// TIA Portal V19 program export: 0 tag tables, 0 data types, 8 data blocks, 41 code blocks (in call order from the OBs), 0 instance data blocks

DATA_BLOCK "ROLL_DB15"   // DB4
{ S7_Optimized_Access := 'TRUE' }
VERSION : 0.1
// stored: AutoNumber true, DBAccessibleFromOPCUA true, DBAccessibleFromWebserver true, IsOnlyStoredInLoadMemory false, IsRetainMemResEnabled false, IsWriteProtectedInAS false, MemoryReserve 100
   VAR RETAIN
      DW : Array[0..131] of Word;
   END_VAR
BEGIN
   DW[0..16] := WORD#16#FFFF;
   DW[17] := WORD#16#3360;
   DW[18..23] := WORD#16#FFFF;
   DW[24] := WORD#16#1010;
   DW[25] := WORD#16#1020;
   DW[26..30] := WORD#16#FFFF;
   DW[31..32] := WORD#16#3120;
   DW[33] := WORD#16#2900;
   DW[34..52] := WORD#16#FFFF;
   DW[53..54] := WORD#16#2120;
   DW[55] := WORD#16#1010;
   DW[56] := WORD#16#2060;
   DW[57] := WORD#16#FFFF;
   DW[58..59] := WORD#16#3180;
   DW[60] := WORD#16#2060;
   DW[61..62] := WORD#16#2600;
   DW[63] := WORD#16#2010;
   DW[64] := WORD#16#FFFF;
   DW[65] := WORD#16#2015;
   DW[66] := WORD#16#FFFF;
   DW[67] := WORD#16#1050;
   DW[68..74] := WORD#16#FFFF;
   DW[75] := WORD#16#2600;
   DW[76] := WORD#16#FFFF;
   DW[77] := WORD#16#2300;
   DW[78..84] := WORD#16#FFFF;
   DW[85] := WORD#16#2120;
   DW[86..101] := WORD#16#FFFF;
   DW[102..103] := WORD#16#2300;
   DW[104..105] := WORD#16#FFFF;
   DW[106] := WORD#16#2010;
   DW[107] := WORD#16#2015;
   DW[108..114] := WORD#16#FFFF;
   DW[115..117] := WORD#16#1050;
   DW[118..126] := WORD#16#FFFF;
   DW[127] := WORD#16#0038;
   DW[128..129] := WORD#16#0011;
   DW[130] := WORD#16#3360;
END_DATA_BLOCK

DATA_BLOCK "ROLL_DB19"   // DB5
{ S7_Optimized_Access := 'TRUE' }
VERSION : 0.1
// stored: AutoNumber true, DBAccessibleFromOPCUA true, DBAccessibleFromWebserver true, IsOnlyStoredInLoadMemory false, IsRetainMemResEnabled false, IsWriteProtectedInAS false, MemoryReserve 100
   VAR RETAIN
      DW : Array[0..131] of Word;
   END_VAR
BEGIN
   DW[0] := WORD#16#FFFF;
   DW[1] := WORD#16#0020;
   DW[2] := WORD#16#0014;
   DW[3..127] := WORD#16#FFFF;
   DW[128..129] := WORD#16#0001;
   DW[130] := WORD#16#0020;
END_DATA_BLOCK

DATA_BLOCK "ROLL_DB205"   // DB8
{ S7_Optimized_Access := 'TRUE' }
VERSION : 0.1
// stored: AutoNumber true, DBAccessibleFromOPCUA true, DBAccessibleFromWebserver true, IsOnlyStoredInLoadMemory false, IsRetainMemResEnabled false, IsWriteProtectedInAS false, MemoryReserve 100
   VAR RETAIN
      DW : Array[0..41] of Word;
   END_VAR
BEGIN
   DW[5] := WORD#16#2360;
   DW[9] := WORD#16#2090;
   DW[13] := WORD#16#0001;
   DW[17] := WORD#16#2240;
   DW[21] := WORD#16#2060;
   DW[25] := WORD#16#2300;
   DW[29] := WORD#16#2120;
   DW[33] := WORD#16#2400;
   DW[37] := WORD#16#0001;
END_DATA_BLOCK

DATA_BLOCK "ROLL_HMI"   // DB3
{ S7_Optimized_Access := 'TRUE' }
VERSION : 0.1
// Flat, symbolic WinCC interface; TP900 control binding is a separate build step.
// stored: AutoNumber true, DBAccessibleFromOPCUA true, DBAccessibleFromWebserver true, IsOnlyStoredInLoadMemory false, IsRetainMemResEnabled false, IsWriteProtectedInAS false, MemoryReserve 100
   VAR
      Heartbeat : DInt;
      Connected : Bool;
      ManualFunction : Int := 255;
      GroundHeld : Bool;
      WorkHeld : Bool;
      KeyF : Array[1..16] of Bool;
      SelectedProgram : Int := 1;
      RecipeCommand : Int := 1;
      RecipeRequest : DInt;
      RecipeAck : DInt;
      RecipeError : Int;
      CurrentProgram : Int := 1;
      ParameterRequest : DInt;
      ParameterAck : DInt;
      ParameterDb : Int := 15;
      ParameterIndex : Int;
      ParameterValue : DInt;
      ParameterCurrentValue : DInt;
      ParameterSlotPresent : Bool;
      ParameterError : Int;
      Dwell1Seconds : Int := 360;
      Drain1Seconds : Int := 90;
      Ultrasound1 : Bool := TRUE;
      Dwell2Seconds : Int := 240;
      Drain2Seconds : Int := 60;
      Dwell3Seconds : Int := 300;
      Drain3Seconds : Int := 120;
      Dry4Seconds : Int := 400;
      BasketMotion : Int := 1;
      BathLift : Bool;
      ProcessTimer1Units : Int;
      ProcessTimer2Units : Int;
      StatusM : Array[0..255, 0..7] of Bool;
      LogicalOutputs : Array[16..25, 0..7] of Bool;
   END_VAR
BEGIN
END_DATA_BLOCK

DATA_BLOCK "ROLL_IO"   // DB2
{ S7_Optimized_Access := 'TRUE' }
VERSION : 0.1
// stored: AutoNumber true, DBAccessibleFromOPCUA true, DBAccessibleFromWebserver true, IsOnlyStoredInLoadMemory false, IsRetainMemResEnabled false, IsWriteProtectedInAS false, MemoryReserve 100
   VAR
      Input : Array[0..127, 0..7] of Bool;
      Output : Array[0..127, 0..7] of Bool;
      Simulation : Bool := TRUE;
      PhysicalOutputsEnabled : Bool := FALSE;
      PhysicalIoConfigured : Bool := FALSE;
      ConversionFault : Bool;
      FirstCycle : Bool := TRUE;
      RuntimeMemory : LReal;
      ClockMs : LReal;
      HmiElapsedMs : LReal;
      HmiLastHeartbeat : DInt;
   END_VAR
BEGIN
END_DATA_BLOCK

DATA_BLOCK "ROLL_Recipe1"   // DB6
{ S7_Optimized_Access := 'TRUE' }
VERSION : 0.1
// stored: AutoNumber true, DBAccessibleFromOPCUA true, DBAccessibleFromWebserver true, IsOnlyStoredInLoadMemory false, IsRetainMemResEnabled false, IsWriteProtectedInAS false, MemoryReserve 100
   VAR RETAIN
      DW : Array[0..41] of Word;
   END_VAR
BEGIN
   DW[5] := WORD#16#2360;
   DW[9] := WORD#16#2090;
   DW[13] := WORD#16#0001;
   DW[17] := WORD#16#2240;
   DW[21] := WORD#16#2060;
   DW[25] := WORD#16#2300;
   DW[29] := WORD#16#2120;
   DW[33] := WORD#16#2400;
   DW[37] := WORD#16#0001;
END_DATA_BLOCK

DATA_BLOCK "ROLL_Recipe2"   // DB7
{ S7_Optimized_Access := 'TRUE' }
VERSION : 0.1
// stored: AutoNumber true, DBAccessibleFromOPCUA true, DBAccessibleFromWebserver true, IsOnlyStoredInLoadMemory false, IsRetainMemResEnabled false, IsWriteProtectedInAS false, MemoryReserve 100
   VAR RETAIN
      DW : Array[0..41] of Word;
   END_VAR
BEGIN
   DW[5] := WORD#16#2360;
   DW[9] := WORD#16#2090;
   DW[13] := WORD#16#0001;
   DW[17] := WORD#16#2240;
   DW[21] := WORD#16#2060;
   DW[25] := WORD#16#2300;
   DW[29] := WORD#16#2120;
   DW[33] := WORD#16#2400;
   DW[37] := WORD#16#0001;
END_DATA_BLOCK

DATA_BLOCK "ROLL_State"   // DB1
{ S7_Optimized_Access := 'TRUE' }
VERSION : 0.1
// stored: AutoNumber true, DBAccessibleFromOPCUA true, DBAccessibleFromWebserver true, IsOnlyStoredInLoadMemory false, IsRetainMemResEnabled false, IsWriteProtectedInAS false, MemoryReserve 100
   VAR RETAIN
      "M" : Array[0..255, 0..7] of Bool;
      S5Timers { S7_SetPoint := 'True'} : Array[0..127] of "ROLL_TimerState";
      S5Counters { S7_SetPoint := 'True'} : Array[0..127] of "ROLL_CounterState";
      CurrentProgram : Int := 1;
   END_VAR
BEGIN
   "M"[0,4] := TRUE;
END_DATA_BLOCK

ORGANIZATION_BLOCK "OB1"   // OB1, SCL, ProgramCycle
TITLE = "Main Program Sweep (Cycle)"
{ S7_Optimized_Access := 'TRUE' }
VERSION : 0.1
// stored: AutoNumber true, IsIECCheckEnabled false, SetENOAutomatically false
   VAR_INPUT
      Initial_Call : Bool;   // Initial call of this OB
      Remanence : Bool;   // =True, if remanent data are available
   END_VAR
BEGIN

   "ROLL_Cycle"();
END_ORGANIZATION_BLOCK

ORGANIZATION_BLOCK "OB100"   // OB100, SCL, Startup
TITLE = "Complete Restart"
{ S7_Optimized_Access := 'TRUE' }
VERSION : 0.1
// stored: AutoNumber true, IsIECCheckEnabled false, SetENOAutomatically false
   VAR_INPUT
      LostRetentive : Bool;   // True if retentive data are lost
      LostRTC : Bool;   // True if date and time are lost
   END_VAR
   VAR_TEMP
      n : Int;
   END_VAR
BEGIN

   // RE plus RS120 bit 3: all M retained. Default T/Z 0..63 retained.
   FOR #n := 64 TO 127 DO
       "ROLL_State".S5Timers[#n].RemainingMs := 0.0;
       "ROLL_State".S5Timers[#n].BaseMs := 0;
       "ROLL_State".S5Timers[#n].Mode := 0;
       "ROLL_State".S5Timers[#n].Q := FALSE;
       "ROLL_State".S5Timers[#n].Previous := FALSE;
       "ROLL_State".S5Counters[#n].Value := 0;
       "ROLL_State".S5Counters[#n].SetPrevious := FALSE;
       "ROLL_State".S5Counters[#n].UpPrevious := FALSE;
       "ROLL_State".S5Counters[#n].DownPrevious := FALSE;
   END_FOR;
   "ROLL_IO".FirstCycle := TRUE;
   "ROLL_IO".ClockMs := 0.0;
   "ROLL_IO".RuntimeMemory := 0.0;
   "ROLL_IO".PhysicalOutputsEnabled := FALSE;
   "ROLL_HMI".Connected := FALSE;
   "ROLL_State".M[0, 1] := TRUE;
   "ROLL_State".M[0, 2] := TRUE;
   "ROLL_State".M[191, 0] := TRUE;
   "ROLL_State".M[190, 5] := FALSE;
   "ROLL_State".M[190, 6] := FALSE;
   "ROLL_State".M[190, 1] := TRUE;
   "ROLL_State".M[191, 4] := TRUE;
   "ROLL_FB90"();
   "ROLL_ShowRecipe"();
END_ORGANIZATION_BLOCK

FUNCTION "ROLL_AdvanceTime" : Void   // FC9, SCL
{ S7_Optimized_Access := 'TRUE' }
VERSION : 0.1
// stored: AutoNumber true, IsIECCheckEnabled false, SetENOAutomatically false, UDAEnableTagReadback false
   VAR_INPUT
      DeltaMs : LReal;
   END_VAR
   VAR_TEMP
      n : Int;
   END_VAR
BEGIN

   IF #DeltaMs < 0.0 THEN
       "ROLL_IO".ConversionFault := TRUE;
       RETURN;
   END_IF;
   FOR #n := 0 TO 127 DO
       IF "ROLL_State".S5Timers[#n].RemainingMs > 0.0 THEN
           "ROLL_State".S5Timers[#n].RemainingMs := "ROLL_State".S5Timers[#n].RemainingMs - #DeltaMs;
           IF "ROLL_State".S5Timers[#n].RemainingMs <= 0.0 THEN
               "ROLL_State".S5Timers[#n].RemainingMs := 0.0;
               "ROLL_State".S5Timers[#n].Q := "ROLL_State".S5Timers[#n].Mode = 0;
           END_IF;
       END_IF;
   END_FOR;
   "ROLL_IO".ClockMs := "ROLL_IO".ClockMs + #DeltaMs;
   WHILE "ROLL_IO".ClockMs >= 250.0 DO
       "ROLL_IO".ClockMs := "ROLL_IO".ClockMs - 250.0;
       "ROLL_State".M[3, 4] := NOT "ROLL_State".M[3, 4];
       IF NOT "ROLL_State".M[3, 4] THEN
           "ROLL_State".M[3, 5] := NOT "ROLL_State".M[3, 5];
           IF NOT "ROLL_State".M[3, 5] THEN
               "ROLL_State".M[3, 6] := NOT "ROLL_State".M[3, 6];
               IF NOT "ROLL_State".M[3, 6] THEN
                   "ROLL_State".M[3, 7] := NOT "ROLL_State".M[3, 7];
               END_IF;
           END_IF;
       END_IF;
   END_WHILE;
END_FUNCTION

FUNCTION "ROLL_CounterOp" : Void   // FC8, SCL
{ S7_Optimized_Access := 'TRUE' }
VERSION : 0.1
// stored: AutoNumber true, IsIECCheckEnabled false, SetENOAutomatically false, UDAEnableTagReadback false
   VAR_INPUT
      Number : Int;
      Operation : Int;   // 0=S set; 1=R reset; 2=ZV up; 3=ZR down
      Signal : Bool;
      Preset : Word;
   END_VAR
   VAR_TEMP
      count : Int;
   END_VAR
BEGIN

   IF (#Number < 0) OR (#Number > 127) THEN
       "ROLL_IO".ConversionFault := TRUE;
       RETURN;
   END_IF;
   CASE #Operation OF
       0:
           IF #Signal AND NOT "ROLL_State".S5Counters[#Number].SetPrevious THEN
               #count := "ROLL_DecodeBCD"(Value := #Preset);
               IF #count >= 0 THEN
                   "ROLL_State".S5Counters[#Number].Value := #count;
               END_IF;
           END_IF;
           "ROLL_State".S5Counters[#Number].SetPrevious := #Signal;
       1:
           IF #Signal THEN
               "ROLL_State".S5Counters[#Number].Value := 0;
           END_IF;
       2:
           IF #Signal AND NOT "ROLL_State".S5Counters[#Number].UpPrevious AND ("ROLL_State".S5Counters[#Number].Value < 999) THEN
               "ROLL_State".S5Counters[#Number].Value := "ROLL_State".S5Counters[#Number].Value + 1;
           END_IF;
           "ROLL_State".S5Counters[#Number].UpPrevious := #Signal;
       3:
           IF #Signal AND NOT "ROLL_State".S5Counters[#Number].DownPrevious AND ("ROLL_State".S5Counters[#Number].Value > 0) THEN
               "ROLL_State".S5Counters[#Number].Value := "ROLL_State".S5Counters[#Number].Value - 1;
           END_IF;
           "ROLL_State".S5Counters[#Number].DownPrevious := #Signal;
       ELSE
           "ROLL_IO".ConversionFault := TRUE;
   END_CASE;
END_FUNCTION

FUNCTION "ROLL_Cycle" : Void   // FC39, SCL
{ S7_Optimized_Access := 'TRUE' }
VERSION : 0.1
// stored: AutoNumber true, IsIECCheckEnabled false, SetENOAutomatically false, UDAEnableTagReadback false
   VAR_TEMP
      delta : LReal;
   END_VAR
BEGIN

   #delta := RUNTIME("ROLL_IO".RuntimeMemory) * 1000.0;
   IF "ROLL_IO".FirstCycle THEN
       #delta := 0.0;
       "ROLL_IO".FirstCycle := FALSE;
   END_IF;
   "ROLL_ReadInputs"();
   "ROLL_AdvanceTime"(DeltaMs := #delta);
   // Exact OB1 order for the process blocks; startup DB creation is replaced.
   IF NOT "ROLL_State".M[0, 2] THEN
       "ROLL_State".M[0, 1] := FALSE;
   END_IF;
   IF "ROLL_State".M[0, 1] THEN
       "ROLL_State".M[0, 7] := TRUE;
   END_IF;
   "ROLL_State".M[0, 5] := NOT "ROLL_State".M[0, 5];
   IF "ROLL_State".M[3, 2] THEN
       "ROLL_State".M[3, 3] := TRUE;
   END_IF;
   IF "ROLL_IO".Input[0, 2] THEN
       "ROLL_State".M[3, 3] := FALSE;
   END_IF;
   "ROLL_State".M[3, 2] := "ROLL_IO".Input[0, 1] AND NOT "ROLL_State".M[0, 1];
   "ROLL_PB2"();
   IF "ROLL_State".M[0, 7] THEN
       "ROLL_State".M[0, 7] := FALSE;
   END_IF;
   "ROLL_PB3"();
   "ROLL_PB4"();
   "ROLL_PB19"();
   "ROLL_PB21"();
   "ROLL_PB50"();
   "ROLL_PB51"();
   "ROLL_PB52"();
   IF NOT "ROLL_State".M[3, 3] THEN
       "ROLL_PB8"();
   END_IF;
   IF NOT "ROLL_State".M[3, 3] THEN
       "ROLL_PB9"();
   END_IF;
   IF NOT "ROLL_State".M[3, 3] THEN
       "ROLL_PB10"();
   END_IF;
   IF NOT "ROLL_State".M[3, 3] THEN
       "ROLL_PB14"();
   END_IF;
   IF "ROLL_State".M[3, 3] THEN
       "ROLL_PB16"();
   END_IF;
   "ROLL_PB7"();
   "ROLL_PB13"();
   "ROLL_PB15"();
   "ROLL_PB17"();
   "ROLL_PB20"();
   "ROLL_PB23"();
   "ROLL_PB24"();
   "ROLL_PB25"();
   "ROLL_FB111"();
   "ROLL_HmiExchange"(DeltaMs := #delta);
   "ROLL_WriteOutputs"();
END_FUNCTION

FUNCTION "ROLL_DecodeBCD" : Int   // FC4, SCL
{ S7_Optimized_Access := 'TRUE' }
VERSION : 0.1
// stored: AutoNumber true, IsIECCheckEnabled false, SetENOAutomatically false, UDAEnableTagReadback false
   VAR_INPUT
      Value : Word;
   END_VAR
   VAR_TEMP
      hundreds : Int;
      tens : Int;
      units : Int;
   END_VAR
BEGIN

   #hundreds := WORD_TO_INT(SHR(IN := #Value AND W#16#0F00, N := 8));
   #tens := WORD_TO_INT(SHR(IN := #Value AND W#16#00F0, N := 4));
   #units := WORD_TO_INT(#Value AND W#16#000F);
   IF (#hundreds > 9) OR (#tens > 9) OR (#units > 9) THEN
       "ROLL_IO".ConversionFault := TRUE;
       #ROLL_DecodeBCD := -1;
   ELSE
       #ROLL_DecodeBCD := #hundreds * 100 + #tens * 10 + #units;
   END_IF;
END_FUNCTION

FUNCTION "ROLL_EncodeSeconds" : Word   // FC5, SCL
{ S7_Optimized_Access := 'TRUE' }
VERSION : 0.1
// stored: AutoNumber true, IsIECCheckEnabled false, SetENOAutomatically false, UDAEnableTagReadback false
   VAR_INPUT
      Seconds : Int;
   END_VAR
BEGIN

   IF (#Seconds < 0) OR (#Seconds > 999) THEN
       #ROLL_EncodeSeconds := W#16#FFFF;
   ELSE
       #ROLL_EncodeSeconds := W#16#2000 OR SHL(IN := INT_TO_WORD(#Seconds / 100), N := 8)
       OR SHL(IN := INT_TO_WORD((#Seconds / 10) MOD 10), N := 4) OR INT_TO_WORD(#Seconds MOD 10);
   END_IF;
END_FUNCTION

FUNCTION "ROLL_FB111" : Void   // FC13, SCL
{ S7_Optimized_Access := 'TRUE' }
VERSION : 0.1
// stored: AutoNumber true, IsIECCheckEnabled false, SetENOAutomatically false, UDAEnableTagReadback false
   VAR_TEMP
      preset : Word;
      signal : Bool;
   END_VAR
BEGIN

   #preset := W#16#2010;
   IF "ROLL_State".M[40, 5] THEN
       #preset := "ROLL_DB205".DW[5];
   ELSIF "ROLL_State".M[42, 1] THEN
       #preset := "ROLL_DB205".DW[17];
   ELSIF "ROLL_State".M[43, 5] THEN
       #preset := "ROLL_DB205".DW[25];
   ELSIF "ROLL_State".M[45, 2] THEN
       #preset := "ROLL_DB205".DW[33];
   END_IF;
   #signal := "ROLL_State".M[40, 5] OR "ROLL_State".M[42, 1] OR "ROLL_State".M[43, 5] OR "ROLL_State".M[45, 2]
   OR "ROLL_State".M[46, 5] OR "ROLL_State".M[48, 1] OR "ROLL_State".M[49, 5] OR "ROLL_State".M[51, 1];
   "ROLL_TimerOp"(Number := 1,
                  Operation := 0,
                  Signal := #signal,
                  Preset := #preset);
   IF (WORD_TO_INT("ROLL_TimerValue"(Number := 1)) <= 7)
       AND ("ROLL_State".M[40, 5] OR "ROLL_State".M[42, 1] OR "ROLL_State".M[43, 5]) AND "ROLL_State".M[111, 5] THEN
       "ROLL_State".M[58, 5] := TRUE;
   END_IF;
   IF "ROLL_State".M[63, 1] AND "ROLL_IO".Input[13, 3] THEN
       "ROLL_State".M[58, 5] := FALSE;
   END_IF;
   #preset := W#16#2010;
   IF "ROLL_State".M[41, 1] THEN
       #preset := "ROLL_DB205".DW[9];
   ELSIF "ROLL_State".M[42, 5] THEN
       #preset := "ROLL_DB205".DW[21];
   ELSIF "ROLL_State".M[44, 1] THEN
       #preset := "ROLL_DB205".DW[29];
   END_IF;
   #signal := "ROLL_State".M[41, 1] OR "ROLL_State".M[42, 5] OR "ROLL_State".M[44, 1]
   OR "ROLL_State".M[45, 6] OR "ROLL_State".M[47, 1] OR "ROLL_State".M[48, 5] OR "ROLL_State".M[50, 1];
   "ROLL_TimerOp"(Number := 2,
                  Operation := 0,
                  Signal := #signal,
                  Preset := #preset);
END_FUNCTION

FUNCTION "ROLL_FB69" : Void   // FC10, SCL
{ S7_Optimized_Access := 'TRUE' }
VERSION : 0.1
// stored: AutoNumber true, IsIECCheckEnabled false, SetENOAutomatically false, UDAEnableTagReadback false
BEGIN

   IF "ROLL_State".M[240, 0] AND "ROLL_State".M[240, 1] THEN
       "ROLL_SetMWord"(FirstByte := 240,
                       Value := W#16#2005);
   ELSE
       "ROLL_SetMWord"(FirstByte := 240,
                       Value := W#16#1005);
   END_IF;
END_FUNCTION

FUNCTION "ROLL_FB90" : Void   // FC12, SCL
{ S7_Optimized_Access := 'TRUE' }
VERSION : 0.1
// stored: AutoNumber true, IsIECCheckEnabled false, SetENOAutomatically false, UDAEnableTagReadback false
BEGIN

   "ROLL_State".M[110, 0] := ("ROLL_DB205".DW[5] AND W#16#0FFF) <> W#16#0000;
   "ROLL_State".M[110, 1] := ("ROLL_DB205".DW[17] AND W#16#0FFF) <> W#16#0000;
   "ROLL_State".M[110, 2] := ("ROLL_DB205".DW[25] AND W#16#0FFF) <> W#16#0000;
   "ROLL_State".M[110, 3] := ("ROLL_DB205".DW[33] AND W#16#0FFF) <> W#16#0000;
   "ROLL_State".M[111, 0] := "ROLL_DB205".DW[37] = W#16#0001;
   "ROLL_State".M[111, 1] := "ROLL_DB205".DW[37] = W#16#0002;
   "ROLL_State".M[111, 2] := "ROLL_DB205".DW[37] = W#16#0003;
   "ROLL_State".M[111, 5] := "ROLL_DB205".DW[37] = W#16#0004;
   "ROLL_State".M[111, 3] := "ROLL_DB205".DW[41] = W#16#0001;
   "ROLL_State".M[111, 4] := "ROLL_DB205".DW[13] = W#16#0001;
   "ROLL_SetMWord"(FirstByte := 250,
                   Value := W#16#0000);
END_FUNCTION

FUNCTION "ROLL_GetDW" : Word   // FC3, SCL
{ S7_Optimized_Access := 'TRUE' }
VERSION : 0.1
// stored: AutoNumber true, IsIECCheckEnabled false, SetENOAutomatically false, UDAEnableTagReadback false
   VAR_INPUT
      DbNumber : Int;
      Index : Int;
   END_VAR
BEGIN

   #ROLL_GetDW := W#16#0000;
   IF (#Index < 0) OR (#Index > 131) THEN
       "ROLL_IO".ConversionFault := TRUE;
       RETURN;
   END_IF;
   CASE #DbNumber OF
       15:
           #ROLL_GetDW := "ROLL_DB15".DW[#Index];
       19:
           #ROLL_GetDW := "ROLL_DB19".DW[#Index];
       ELSE
           "ROLL_IO".ConversionFault := TRUE;
   END_CASE;
END_FUNCTION

FUNCTION "ROLL_GetM" : Word   // FC1, SCL
{ S7_Optimized_Access := 'TRUE' }
VERSION : 0.1
// stored: AutoNumber true, IsIECCheckEnabled false, SetENOAutomatically false, UDAEnableTagReadback false
   VAR_INPUT
      FirstByte : Int;
      Width : Int;
   END_VAR
   VAR_TEMP
      "b" : Int;
      n : Int;
      bit : Int;
      mask : Word;
      result : Word;
   END_VAR
BEGIN

   #result := W#16#0000;
   IF (#FirstByte < 0) OR (#FirstByte > 255) OR ((#Width <> 8) AND (#Width <> 16)) OR ((#Width = 16) AND (#FirstByte > 254)) THEN
       "ROLL_IO".ConversionFault := TRUE;
       #ROLL_GetM := #result;
       RETURN;
   END_IF;
   FOR #n := 0 TO (#Width / 8) - 1 DO
       #b := #FirstByte + #n;
       FOR #bit := 0 TO 7 DO
           #mask := SHL(IN := W#16#0001, N := #bit + (#Width - 8 - 8 * #n));
           IF "ROLL_State".M[#b, #bit] THEN
               #result := #result OR #mask;
           END_IF;
       END_FOR;
   END_FOR;
   #ROLL_GetM := #result;
END_FUNCTION

FUNCTION "ROLL_HmiExchange" : Void   // FC38, SCL
{ S7_Optimized_Access := 'TRUE' }
VERSION : 0.1
// stored: AutoNumber true, IsIECCheckEnabled false, SetENOAutomatically false, UDAEnableTagReadback false
   VAR_INPUT
      DeltaMs : LReal;
   END_VAR
   VAR_TEMP
      "b" : Int;
      bit : Int;
      n : Int;
      fieldIndex : Int;
      index : Int;
      raw : Word;
      base : DInt;
      count : DInt;
      recipe : Array[0..41] of Word;
   END_VAR
BEGIN

   // Called at the end of the scan, like the former OP15 functions in OB1.
   "ROLL_IO".HmiElapsedMs := "ROLL_IO".HmiElapsedMs + #DeltaMs;
   IF "ROLL_HMI".Heartbeat <> "ROLL_IO".HmiLastHeartbeat THEN
       "ROLL_IO".HmiLastHeartbeat := "ROLL_HMI".Heartbeat;
       "ROLL_IO".HmiElapsedMs := 0.0;
       "ROLL_HMI".Connected := TRUE;
   END_IF;
   IF "ROLL_IO".HmiElapsedMs >= 1500.0 THEN
       "ROLL_HMI".Connected := FALSE;
   END_IF;
   "ROLL_State".M[190, 5] := "ROLL_HMI".Connected AND "ROLL_HMI".GroundHeld;
   "ROLL_State".M[190, 6] := "ROLL_HMI".Connected AND "ROLL_HMI".WorkHeld;
   "ROLL_State".M[190, 3] := ("ROLL_State".M[190, 5] OR "ROLL_State".M[190, 6]) AND NOT "ROLL_State".M[190, 4];
   "ROLL_State".M[190, 4] := "ROLL_State".M[190, 5] OR "ROLL_State".M[190, 6];
   "ROLL_State".M[191, 0] := FALSE;
   IF ("ROLL_HMI".ManualFunction >= 0) AND ("ROLL_HMI".ManualFunction <= 255) AND "ROLL_HMI".Connected THEN
       "ROLL_SetMWord"(FirstByte := 238,
                       Value := INT_TO_WORD("ROLL_HMI".ManualFunction));
   ELSE
       "ROLL_SetMWord"(FirstByte := 238,
                       Value := W#16#00FF);
   END_IF;
   FOR #n := 0 TO 7 DO
       "ROLL_State".M[192, #n] := "ROLL_HMI".Connected AND "ROLL_HMI".KeyF[#n + 1];
       "ROLL_State".M[193, #n] := "ROLL_HMI".Connected AND "ROLL_HMI".KeyF[#n + 9];
   END_FOR;

   // Request/acknowledgement counters prevent partial edits on every scan.
   // Command 1 loads the retained program; command 2 saves the displayed values.
   IF "ROLL_HMI".RecipeRequest <> "ROLL_HMI".RecipeAck THEN
       "ROLL_HMI".RecipeError := 0;
       IF NOT "ROLL_HMI".Connected THEN
           "ROLL_HMI".RecipeError := 8;
       ELSIF ("ROLL_HMI".SelectedProgram < 1) OR ("ROLL_HMI".SelectedProgram > 2) THEN
           "ROLL_HMI".RecipeError := 1;
       ELSIF NOT "ROLL_IO".Input[0, 1] THEN
           "ROLL_HMI".RecipeError := 2; // requires manual operating mode
       ELSIF ("ROLL_HMI".RecipeCommand <> 1) AND ("ROLL_HMI".RecipeCommand <> 2) THEN
           "ROLL_HMI".RecipeError := 3;
       ELSE
           FOR #n := 0 TO 41 DO
               IF "ROLL_HMI".SelectedProgram = 1 THEN
                   #recipe[#n] := "ROLL_Recipe1".DW[#n];
               ELSE
                   #recipe[#n] := "ROLL_Recipe2".DW[#n];
               END_IF;
           END_FOR;
           IF "ROLL_HMI".RecipeCommand = 2 THEN
               #recipe[5] := "ROLL_EncodeSeconds"(Seconds := "ROLL_HMI".Dwell1Seconds);
               #recipe[9] := "ROLL_EncodeSeconds"(Seconds := "ROLL_HMI".Drain1Seconds);
               #recipe[17] := "ROLL_EncodeSeconds"(Seconds := "ROLL_HMI".Dwell2Seconds);
               #recipe[21] := "ROLL_EncodeSeconds"(Seconds := "ROLL_HMI".Drain2Seconds);
               #recipe[25] := "ROLL_EncodeSeconds"(Seconds := "ROLL_HMI".Dwell3Seconds);
               #recipe[29] := "ROLL_EncodeSeconds"(Seconds := "ROLL_HMI".Drain3Seconds);
               #recipe[33] := "ROLL_EncodeSeconds"(Seconds := "ROLL_HMI".Dry4Seconds);
               FOR #n := 0 TO 6 DO
                   CASE #n OF
                       0:
                           #fieldIndex := 5;
                       1:
                           #fieldIndex := 9;
                       2:
                           #fieldIndex := 17;
                       3:
                           #fieldIndex := 21;
                       4:
                           #fieldIndex := 25;
                       5:
                           #fieldIndex := 29;
                       6:
                           #fieldIndex := 33;
                   END_CASE;
                   IF #recipe[#fieldIndex] = W#16#FFFF THEN
                       "ROLL_HMI".RecipeError := 4;
                   END_IF;
               END_FOR;
               IF ("ROLL_HMI".BasketMotion < 0) OR ("ROLL_HMI".BasketMotion > 4) THEN
                   "ROLL_HMI".RecipeError := 5;
               END_IF;
               #recipe[37] := INT_TO_WORD("ROLL_HMI".BasketMotion);
               #recipe[13] := W#16#0000;
               IF "ROLL_HMI".Ultrasound1 THEN
                   #recipe[13] := W#16#0001;
               END_IF;
               #recipe[41] := W#16#0000;
               IF "ROLL_HMI".BathLift THEN
                   #recipe[41] := W#16#0001;
               END_IF;
           END_IF;
           IF "ROLL_HMI".RecipeError = 0 THEN
               FOR #n := 0 TO 41 DO
                   "ROLL_DB205".DW[#n] := #recipe[#n];
                   IF "ROLL_HMI".RecipeCommand = 2 THEN
                       IF "ROLL_HMI".SelectedProgram = 1 THEN
                           "ROLL_Recipe1".DW[#n] := #recipe[#n];
                       ELSE
                           "ROLL_Recipe2".DW[#n] := #recipe[#n];
                       END_IF;
                   END_IF;
               END_FOR;
               "ROLL_State".CurrentProgram := "ROLL_HMI".SelectedProgram;
               "ROLL_ShowRecipe"();
               "ROLL_State".M[190, 1] := TRUE;
               "ROLL_State".M[190, 2] := FALSE;
               "ROLL_State".M[191, 4] := TRUE;
               "ROLL_FB90"();
           END_IF;
       END_IF;
       "ROLL_HMI".RecipeAck := "ROLL_HMI".RecipeRequest;
   END_IF;

   IF "ROLL_HMI".ParameterRequest <> "ROLL_HMI".ParameterAck THEN
       "ROLL_HMI".ParameterError := 0;
       #index := "ROLL_HMI".ParameterIndex;
       #raw := W#16#FFFF;
       IF NOT "ROLL_HMI".Connected THEN
           "ROLL_HMI".ParameterError := 8;
       ELSIF (#index < 0) OR (#index > 127) THEN
           "ROLL_HMI".ParameterError := 1;
       ELSIF NOT "ROLL_IO".Input[0, 1] THEN
           "ROLL_HMI".ParameterError := 2;
       ELSIF ("ROLL_HMI".ParameterDb <> 15) AND ("ROLL_HMI".ParameterDb <> 19) THEN
           "ROLL_HMI".ParameterError := 3;
       ELSE
           #raw := "ROLL_GetDW"(DbNumber := "ROLL_HMI".ParameterDb, Index := #index);
           IF #raw = W#16#FFFF THEN
               "ROLL_HMI".ParameterError := 4;
           ELSE
               #base := 1;
               IF "ROLL_HMI".ParameterDb = 15 THEN
                   CASE WORD_TO_INT(SHR(IN := #raw AND W#16#F000, N := 12)) OF
                       0:
                           #base := 10;
                       1:
                           #base := 100;
                       2:
                           #base := 1000;
                       3:
                           #base := 10000;
                       ELSE
                           #base := 0;
                   END_CASE;
               END_IF;
               IF #base = 0 THEN
                   "ROLL_HMI".ParameterError := 5;
               ELSIF ("ROLL_HMI".ParameterValue < 0) OR (("ROLL_HMI".ParameterValue MOD #base) <> 0) THEN
                   "ROLL_HMI".ParameterError := 6;
               ELSE
                   #count := "ROLL_HMI".ParameterValue / #base;
                   IF #count > 999 THEN
                       "ROLL_HMI".ParameterError := 7;
                   ELSE
                       #raw := (#raw AND W#16#F000) OR SHL(IN := DINT_TO_WORD(#count / 100), N := 8)
                       OR SHL(IN := DINT_TO_WORD((#count / 10) MOD 10), N := 4) OR DINT_TO_WORD(#count MOD 10);
                       IF "ROLL_HMI".ParameterDb = 15 THEN
                           "ROLL_DB15".DW[#index] := #raw;
                       ELSE
                           "ROLL_DB19".DW[#index] := #raw;
                       END_IF;
                   END_IF;
               END_IF;
           END_IF;
       END_IF;
       "ROLL_HMI".ParameterAck := "ROLL_HMI".ParameterRequest;
   END_IF;
   "ROLL_HMI".ParameterSlotPresent := FALSE;
   "ROLL_HMI".ParameterCurrentValue := 0;
   #index := "ROLL_HMI".ParameterIndex;
   IF (#index >= 0) AND (#index <= 127) AND (("ROLL_HMI".ParameterDb = 15) OR ("ROLL_HMI".ParameterDb = 19)) THEN
       #raw := "ROLL_GetDW"(DbNumber := "ROLL_HMI".ParameterDb, Index := #index);
       IF #raw <> W#16#FFFF THEN
           #count := INT_TO_DINT("ROLL_DecodeBCD"(Value := #raw));
           #base := 1;
           IF "ROLL_HMI".ParameterDb = 15 THEN
               CASE WORD_TO_INT(SHR(IN := #raw AND W#16#F000, N := 12)) OF
                   0:
                       #base := 10;
                   1:
                       #base := 100;
                   2:
                       #base := 1000;
                   3:
                       #base := 10000;
                   ELSE
                       #base := 0;
               END_CASE;
           END_IF;
           IF (#count >= 0) AND (#base > 0) THEN
               "ROLL_HMI".ParameterSlotPresent := TRUE;
               "ROLL_HMI".ParameterCurrentValue := #count * #base;
           END_IF;
       END_IF;
   END_IF;
   IF WORD_TO_INT("ROLL_GetM"(FirstByte := 239, Width := 8)) <> 255 THEN
       "ROLL_PB18"();
   ELSE
       "ROLL_SetMWord"(FirstByte := 250,
                       Value := W#16#0000);
       "ROLL_SetMWord"(FirstByte := 252,
                       Value := W#16#0000);
   END_IF;
   "ROLL_HMI".ProcessTimer1Units := WORD_TO_INT("ROLL_TimerValue"(Number := 1));
   "ROLL_HMI".ProcessTimer2Units := WORD_TO_INT("ROLL_TimerValue"(Number := 2));
   FOR #b := 0 TO 255 DO
       FOR #bit := 0 TO 7 DO
           "ROLL_HMI".StatusM[#b, #bit] := "ROLL_State".M[#b, #bit];
       END_FOR;
   END_FOR;
   FOR #b := 16 TO 25 DO
       FOR #bit := 0 TO 7 DO
           "ROLL_HMI".LogicalOutputs[#b, #bit] := "ROLL_IO".Output[#b, #bit];
       END_FOR;
   END_FOR;
END_FUNCTION

FUNCTION "ROLL_PB10" : Void   // FC20, SCL
{ S7_Optimized_Access := 'TRUE' }
VERSION : 0.1
// stored: AutoNumber true, IsIECCheckEnabled false, SetENOAutomatically false, UDAEnableTagReadback false
   VAR_TEMP
      r : Bool;
      a1 : Word;
      a2 : Word;
      activeDataBlock : Int;
      comparisonResults : Array[0..0] of Bool;
   END_VAR
BEGIN

   #r := FALSE;
   #a1 := W#16#0000;
   #a2 := W#16#0000;
   #activeDataBlock := 0;
   // PB10, STEP 5 network 1
   #r := (((NOT "ROLL_State".M[110, 0]) AND (NOT "ROLL_State".M[110, 1]) AND (NOT "ROLL_State".M[110, 2]) AND (NOT "ROLL_State".M[110, 3]) AND "ROLL_State".M[40, 1]) OR ((NOT "ROLL_State".M[110, 1]) AND (NOT "ROLL_State".M[110, 2]) AND (NOT "ROLL_State".M[110, 3]) AND "ROLL_State".M[41, 2]) OR ((NOT "ROLL_State".M[110, 2]) AND (NOT "ROLL_State".M[110, 3]) AND "ROLL_State".M[42, 6]) OR ((NOT "ROLL_State".M[110, 3]) AND "ROLL_State".M[44, 2]) OR "ROLL_State".M[45, 7]);
   "ROLL_State".M[240, 0] := #r;
   // PB10, STEP 5 network 2
   #r := ((NOT "ROLL_IO".Input[119, 6]) AND "ROLL_IO".Input[12, 5] AND "ROLL_IO".Input[12, 7] AND "ROLL_State".M[110, 4] AND "ROLL_State".M[240, 0] AND "ROLL_State".M[35, 2]);
   IF #r THEN
       "ROLL_State".M[46, 2] := TRUE;
   END_IF;
   #r := ("ROLL_State".M[32, 2] OR "ROLL_State".M[46, 3]);
   IF #r THEN
       "ROLL_State".M[46, 2] := FALSE;
   END_IF;
   // PB10, STEP 5 network 3
   #r := ("ROLL_IO".Input[11, 6] AND "ROLL_IO".Input[119, 6] AND "ROLL_State".M[35, 2] AND "ROLL_State".M[46, 2]);
   IF #r THEN
       "ROLL_State".M[46, 3] := TRUE;
   END_IF;
   #r := ("ROLL_State".M[32, 2] OR "ROLL_State".M[46, 4]);
   IF #r THEN
       "ROLL_State".M[46, 3] := FALSE;
   END_IF;
   // PB10, STEP 5 network 4
   #r := ((NOT "ROLL_IO".Input[12, 1]) AND "ROLL_IO".Input[12, 5] AND "ROLL_State".M[35, 2] AND "ROLL_State".M[46, 3]);
   IF #r THEN
       "ROLL_State".M[46, 4] := TRUE;
   END_IF;
   #r := ("ROLL_State".M[32, 2] OR "ROLL_State".M[46, 5]);
   IF #r THEN
       "ROLL_State".M[46, 4] := FALSE;
   END_IF;
   // PB10, STEP 5 network 5
   #r := ("ROLL_IO".Input[12, 1] AND "ROLL_IO".Input[12, 7] AND "ROLL_State".M[35, 2] AND "ROLL_State".M[46, 4]);
   IF #r THEN
       "ROLL_State".M[46, 5] := TRUE;
   END_IF;
   #r := ("ROLL_State".M[32, 2] OR "ROLL_State".M[46, 6]);
   IF #r THEN
       "ROLL_State".M[46, 5] := FALSE;
   END_IF;
   // PB10, STEP 5 network 6
   #r := ("ROLL_State".M[35, 2] AND "ROLL_State".M[46, 5] AND "ROLL_State".S5Timers[1].Q);
   IF #r THEN
       "ROLL_State".M[46, 6] := TRUE;
   END_IF;
   #r := ("ROLL_State".M[32, 2] OR "ROLL_State".M[46, 7]);
   IF #r THEN
       "ROLL_State".M[46, 6] := FALSE;
   END_IF;
   // PB10, STEP 5 network 7
   #r := ("ROLL_State".M[35, 2] AND "ROLL_State".M[46, 6]);
   IF #r THEN
       "ROLL_State".M[46, 7] := TRUE;
   END_IF;
   #r := ("ROLL_State".M[32, 2] OR "ROLL_State".M[47, 0]);
   IF #r THEN
       "ROLL_State".M[46, 7] := FALSE;
   END_IF;
   // PB10, STEP 5 network 8
   #r := ((NOT "ROLL_IO".Input[12, 5]) AND "ROLL_State".M[35, 2] AND "ROLL_State".M[46, 7]);
   IF #r THEN
       "ROLL_State".M[47, 0] := TRUE;
   END_IF;
   #r := ("ROLL_State".M[32, 2] OR "ROLL_State".M[47, 1]);
   IF #r THEN
       "ROLL_State".M[47, 0] := FALSE;
   END_IF;
   // PB10, STEP 5 network 9
   #r := ("ROLL_IO".Input[12, 5] AND "ROLL_IO".Input[12, 7] AND "ROLL_State".M[35, 2] AND "ROLL_State".M[47, 0]);
   IF #r THEN
       "ROLL_State".M[47, 1] := TRUE;
   END_IF;
   #r := ("ROLL_State".M[32, 2] OR "ROLL_State".M[47, 2]);
   IF #r THEN
       "ROLL_State".M[47, 1] := FALSE;
   END_IF;
   // PB10, STEP 5 network 10
   #r := ("ROLL_State".M[35, 2] AND "ROLL_State".M[47, 1] AND "ROLL_State".S5Timers[2].Q);
   IF #r THEN
       "ROLL_State".M[47, 2] := TRUE;
   END_IF;
   #r := ("ROLL_State".M[32, 2] OR "ROLL_State".M[47, 3] OR "ROLL_State".M[47, 6]);
   IF #r THEN
       "ROLL_State".M[47, 2] := FALSE;
   END_IF;
   // PB10, STEP 5 network 11
   #r := ((NOT "ROLL_State".M[110, 5]) AND (NOT "ROLL_State".M[110, 6]) AND "ROLL_State".M[35, 2] AND "ROLL_State".M[47, 2]);
   IF #r THEN
       "ROLL_State".M[47, 3] := TRUE;
   END_IF;
   #r := ("ROLL_State".M[32, 2] OR "ROLL_State".M[47, 4]);
   IF #r THEN
       "ROLL_State".M[47, 3] := FALSE;
   END_IF;
   // PB10, STEP 5 network 12
   #r := ("ROLL_IO".Input[13, 3] AND "ROLL_State".M[35, 2] AND "ROLL_State".M[47, 3] AND "ROLL_State".M[63, 1]);
   IF #r THEN
       "ROLL_State".M[47, 4] := TRUE;
   END_IF;
   #r := ("ROLL_State".M[32, 2] OR "ROLL_State".M[50, 6] OR "ROLL_State".M[52, 0]);
   IF #r THEN
       "ROLL_State".M[47, 4] := FALSE;
   END_IF;
   // PB10, STEP 5 network 13
   #r := (((NOT "ROLL_State".M[110, 0]) AND (NOT "ROLL_State".M[110, 1]) AND (NOT "ROLL_State".M[110, 2]) AND (NOT "ROLL_State".M[110, 3]) AND (NOT "ROLL_State".M[110, 4]) AND "ROLL_State".M[40, 1]) OR ((NOT "ROLL_State".M[110, 1]) AND (NOT "ROLL_State".M[110, 2]) AND (NOT "ROLL_State".M[110, 3]) AND (NOT "ROLL_State".M[110, 4]) AND "ROLL_State".M[41, 2]) OR ((NOT "ROLL_State".M[110, 2]) AND (NOT "ROLL_State".M[110, 3]) AND (NOT "ROLL_State".M[110, 4]) AND "ROLL_State".M[42, 6]) OR ((NOT "ROLL_State".M[110, 3]) AND (NOT "ROLL_State".M[110, 4]) AND "ROLL_State".M[44, 2]) OR ((NOT "ROLL_State".M[110, 4]) AND "ROLL_State".M[45, 7]) OR "ROLL_State".M[47, 2]);
   "ROLL_State".M[240, 0] := #r;
   // PB10, STEP 5 network 14
   #r := ((NOT "ROLL_IO".Input[119, 7]) AND "ROLL_IO".Input[12, 5] AND "ROLL_IO".Input[12, 7] AND "ROLL_State".M[110, 5] AND "ROLL_State".M[240, 0] AND "ROLL_State".M[35, 2]);
   IF #r THEN
       "ROLL_State".M[47, 6] := TRUE;
   END_IF;
   #r := ("ROLL_State".M[32, 2] OR "ROLL_State".M[47, 7]);
   IF #r THEN
       "ROLL_State".M[47, 6] := FALSE;
   END_IF;
   // PB10, STEP 5 network 15
   #r := ("ROLL_IO".Input[11, 6] AND "ROLL_IO".Input[119, 7] AND "ROLL_State".M[35, 2] AND "ROLL_State".M[47, 6]);
   IF #r THEN
       "ROLL_State".M[47, 7] := TRUE;
   END_IF;
   #r := ("ROLL_State".M[32, 2] OR "ROLL_State".M[48, 0]);
   IF #r THEN
       "ROLL_State".M[47, 7] := FALSE;
   END_IF;
   // PB10, STEP 5 network 16
   #r := ((NOT "ROLL_IO".Input[12, 1]) AND "ROLL_IO".Input[12, 5] AND "ROLL_State".M[35, 2] AND "ROLL_State".M[47, 7]);
   IF #r THEN
       "ROLL_State".M[48, 0] := TRUE;
   END_IF;
   #r := ("ROLL_State".M[32, 2] OR "ROLL_State".M[48, 1]);
   IF #r THEN
       "ROLL_State".M[48, 0] := FALSE;
   END_IF;
   // PB10, STEP 5 network 17
   #r := ("ROLL_IO".Input[12, 1] AND "ROLL_IO".Input[12, 7] AND "ROLL_State".M[35, 2] AND "ROLL_State".M[48, 0]);
   IF #r THEN
       "ROLL_State".M[48, 1] := TRUE;
   END_IF;
   #r := ("ROLL_State".M[32, 2] OR "ROLL_State".M[48, 2]);
   IF #r THEN
       "ROLL_State".M[48, 1] := FALSE;
   END_IF;
   // PB10, STEP 5 network 18
   #r := ("ROLL_State".M[35, 2] AND "ROLL_State".M[48, 1] AND "ROLL_State".S5Timers[1].Q);
   IF #r THEN
       "ROLL_State".M[48, 2] := TRUE;
   END_IF;
   #r := ("ROLL_State".M[32, 2] OR "ROLL_State".M[48, 3]);
   IF #r THEN
       "ROLL_State".M[48, 2] := FALSE;
   END_IF;
   // PB10, STEP 5 network 19
   #r := ("ROLL_State".M[35, 2] AND "ROLL_State".M[48, 2]);
   IF #r THEN
       "ROLL_State".M[48, 3] := TRUE;
   END_IF;
   #r := ("ROLL_State".M[32, 2] OR "ROLL_State".M[48, 4]);
   IF #r THEN
       "ROLL_State".M[48, 3] := FALSE;
   END_IF;
   // PB10, STEP 5 network 20
   #r := ((NOT "ROLL_IO".Input[12, 5]) AND "ROLL_State".M[35, 2] AND "ROLL_State".M[48, 3]);
   IF #r THEN
       "ROLL_State".M[48, 4] := TRUE;
   END_IF;
   #r := ("ROLL_State".M[32, 2] OR "ROLL_State".M[48, 5]);
   IF #r THEN
       "ROLL_State".M[48, 4] := FALSE;
   END_IF;
   // PB10, STEP 5 network 21
   #r := ("ROLL_IO".Input[12, 5] AND "ROLL_IO".Input[12, 7] AND "ROLL_State".M[35, 2] AND "ROLL_State".M[48, 4]);
   IF #r THEN
       "ROLL_State".M[48, 5] := TRUE;
   END_IF;
   #r := ("ROLL_State".M[32, 2] OR "ROLL_State".M[48, 6]);
   IF #r THEN
       "ROLL_State".M[48, 5] := FALSE;
   END_IF;
   // PB10, STEP 5 network 22
   #r := ("ROLL_State".M[35, 2] AND "ROLL_State".M[48, 5] AND "ROLL_State".S5Timers[2].Q);
   IF #r THEN
       "ROLL_State".M[48, 6] := TRUE;
   END_IF;
   #r := ("ROLL_State".M[32, 2] OR "ROLL_State".M[48, 7] OR "ROLL_State".M[49, 2]);
   IF #r THEN
       "ROLL_State".M[48, 6] := FALSE;
   END_IF;
   // PB10, STEP 5 network 23
   #r := ((NOT "ROLL_State".M[110, 6]) AND "ROLL_State".M[35, 2] AND "ROLL_State".M[48, 6]);
   IF #r THEN
       "ROLL_State".M[48, 7] := TRUE;
   END_IF;
   #r := ("ROLL_State".M[32, 2] OR "ROLL_State".M[49, 0]);
   IF #r THEN
       "ROLL_State".M[48, 7] := FALSE;
   END_IF;
   // PB10, STEP 5 network 24
   #r := ("ROLL_IO".Input[13, 3] AND "ROLL_State".M[35, 2] AND "ROLL_State".M[48, 7] AND "ROLL_State".M[63, 1]);
   IF #r THEN
       "ROLL_State".M[49, 0] := TRUE;
   END_IF;
   #r := ("ROLL_State".M[32, 2] OR "ROLL_State".M[50, 6] OR "ROLL_State".M[52, 0]);
   IF #r THEN
       "ROLL_State".M[49, 0] := FALSE;
   END_IF;
   // PB10, STEP 5 network 25
   #r := (((NOT "ROLL_State".M[110, 0]) AND (NOT "ROLL_State".M[110, 1]) AND (NOT "ROLL_State".M[110, 2]) AND (NOT "ROLL_State".M[110, 3]) AND (NOT "ROLL_State".M[110, 4]) AND (NOT "ROLL_State".M[110, 5]) AND "ROLL_State".M[40, 1]) OR ((NOT "ROLL_State".M[110, 1]) AND (NOT "ROLL_State".M[110, 2]) AND (NOT "ROLL_State".M[110, 3]) AND (NOT "ROLL_State".M[110, 4]) AND (NOT "ROLL_State".M[110, 5]) AND "ROLL_State".M[41, 2]) OR ((NOT "ROLL_State".M[110, 2]) AND (NOT "ROLL_State".M[110, 3]) AND (NOT "ROLL_State".M[110, 4]) AND (NOT "ROLL_State".M[110, 5]) AND "ROLL_State".M[42, 6]) OR ((NOT "ROLL_State".M[110, 3]) AND (NOT "ROLL_State".M[110, 4]) AND (NOT "ROLL_State".M[110, 5]) AND "ROLL_State".M[44, 2]) OR ((NOT "ROLL_State".M[110, 4]) AND (NOT "ROLL_State".M[110, 5]) AND "ROLL_State".M[45, 7]) OR ((NOT "ROLL_State".M[110, 5]) AND "ROLL_State".M[47, 2]) OR "ROLL_State".M[48, 6]);
   "ROLL_State".M[240, 0] := #r;
   // PB10, STEP 5 network 26
   #r := ((NOT "ROLL_IO".Input[120, 0]) AND "ROLL_IO".Input[12, 5] AND "ROLL_IO".Input[12, 7] AND "ROLL_State".M[110, 6] AND "ROLL_State".M[240, 0] AND "ROLL_State".M[35, 2]);
   IF #r THEN
       "ROLL_State".M[49, 2] := TRUE;
   END_IF;
   #r := ("ROLL_State".M[32, 2] OR "ROLL_State".M[49, 3]);
   IF #r THEN
       "ROLL_State".M[49, 2] := FALSE;
   END_IF;
   // PB10, STEP 5 network 27
   #r := ("ROLL_IO".Input[11, 6] AND "ROLL_IO".Input[120, 0] AND "ROLL_State".M[35, 2] AND "ROLL_State".M[49, 2]);
   IF #r THEN
       "ROLL_State".M[49, 3] := TRUE;
   END_IF;
   #r := ("ROLL_State".M[32, 2] OR "ROLL_State".M[49, 4]);
   IF #r THEN
       "ROLL_State".M[49, 3] := FALSE;
   END_IF;
   // PB10, STEP 5 network 28
   #r := ((NOT "ROLL_IO".Input[12, 1]) AND "ROLL_IO".Input[12, 5] AND "ROLL_State".M[35, 2] AND "ROLL_State".M[49, 3]);
   IF #r THEN
       "ROLL_State".M[49, 4] := TRUE;
   END_IF;
   #r := ("ROLL_State".M[32, 2] OR "ROLL_State".M[49, 5]);
   IF #r THEN
       "ROLL_State".M[49, 4] := FALSE;
   END_IF;
   // PB10, STEP 5 network 29
   #r := ("ROLL_IO".Input[12, 1] AND "ROLL_IO".Input[12, 7] AND "ROLL_State".M[35, 2] AND "ROLL_State".M[49, 4]);
   IF #r THEN
       "ROLL_State".M[49, 5] := TRUE;
   END_IF;
   #r := ("ROLL_State".M[32, 2] OR "ROLL_State".M[49, 6]);
   IF #r THEN
       "ROLL_State".M[49, 5] := FALSE;
   END_IF;
   // PB10, STEP 5 network 30
   #r := ("ROLL_State".M[35, 2] AND "ROLL_State".M[49, 5] AND "ROLL_State".S5Timers[1].Q);
   IF #r THEN
       "ROLL_State".M[49, 6] := TRUE;
   END_IF;
   #r := ("ROLL_State".M[32, 2] OR "ROLL_State".M[49, 7]);
   IF #r THEN
       "ROLL_State".M[49, 6] := FALSE;
   END_IF;
   // PB10, STEP 5 network 31
   #r := ("ROLL_State".M[35, 2] AND "ROLL_State".M[49, 6]);
   IF #r THEN
       "ROLL_State".M[49, 7] := TRUE;
   END_IF;
   #r := ("ROLL_State".M[32, 2] OR "ROLL_State".M[50, 0]);
   IF #r THEN
       "ROLL_State".M[49, 7] := FALSE;
   END_IF;
   // PB10, STEP 5 network 32
   #r := ((NOT "ROLL_IO".Input[12, 5]) AND "ROLL_State".M[35, 2] AND "ROLL_State".M[49, 7]);
   IF #r THEN
       "ROLL_State".M[50, 0] := TRUE;
   END_IF;
   #r := ("ROLL_State".M[32, 2] OR "ROLL_State".M[50, 1]);
   IF #r THEN
       "ROLL_State".M[50, 0] := FALSE;
   END_IF;
   // PB10, STEP 5 network 33
   #r := ("ROLL_IO".Input[12, 5] AND "ROLL_IO".Input[12, 7] AND "ROLL_State".M[35, 2] AND "ROLL_State".M[50, 0]);
   IF #r THEN
       "ROLL_State".M[50, 1] := TRUE;
   END_IF;
   #r := ("ROLL_State".M[32, 2] OR "ROLL_State".M[50, 2]);
   IF #r THEN
       "ROLL_State".M[50, 1] := FALSE;
   END_IF;
   // PB10, STEP 5 network 34
   #r := ("ROLL_State".M[35, 2] AND "ROLL_State".M[50, 1] AND "ROLL_State".S5Timers[2].Q);
   IF #r THEN
       "ROLL_State".M[50, 2] := TRUE;
   END_IF;
   #r := ("ROLL_State".M[32, 2] OR "ROLL_State".M[50, 3]);
   IF #r THEN
       "ROLL_State".M[50, 2] := FALSE;
   END_IF;
   // PB10, STEP 5 network 35
   #r := ("ROLL_State".M[35, 2] AND "ROLL_State".M[50, 2]);
   IF #r THEN
       "ROLL_State".M[50, 3] := TRUE;
   END_IF;
   #r := ("ROLL_State".M[32, 2] OR "ROLL_State".M[50, 4]);
   IF #r THEN
       "ROLL_State".M[50, 3] := FALSE;
   END_IF;
   // PB10, STEP 5 network 36
   #r := ("ROLL_IO".Input[13, 3] AND "ROLL_State".M[35, 2] AND "ROLL_State".M[50, 3] AND "ROLL_State".M[63, 1]);
   IF #r THEN
       "ROLL_State".M[50, 4] := TRUE;
   END_IF;
   #r := ("ROLL_State".M[32, 2] OR "ROLL_State".M[50, 6] OR "ROLL_State".M[52, 0]);
   IF #r THEN
       "ROLL_State".M[50, 4] := FALSE;
   END_IF;
   // PB10, STEP 5 network 37
   #r := (((NOT "ROLL_State".M[110, 0]) AND (NOT "ROLL_State".M[110, 1]) AND (NOT "ROLL_State".M[110, 2]) AND (NOT "ROLL_State".M[110, 3]) AND (NOT "ROLL_State".M[110, 4]) AND (NOT "ROLL_State".M[110, 5]) AND (NOT "ROLL_State".M[110, 6]) AND "ROLL_State".M[40, 1]) OR ((NOT "ROLL_State".M[110, 1]) AND (NOT "ROLL_State".M[110, 2]) AND (NOT "ROLL_State".M[110, 3]) AND (NOT "ROLL_State".M[110, 4]) AND (NOT "ROLL_State".M[110, 5]) AND (NOT "ROLL_State".M[110, 6]) AND "ROLL_State".M[41, 4]) OR ((NOT "ROLL_State".M[110, 2]) AND (NOT "ROLL_State".M[110, 3]) AND (NOT "ROLL_State".M[110, 4]) AND (NOT "ROLL_State".M[110, 5]) AND (NOT "ROLL_State".M[110, 6]) AND "ROLL_State".M[43, 0]));
   "ROLL_State".M[240, 0] := #r;
   // PB10, STEP 5 network 38
   #r := (((NOT "ROLL_State".M[110, 3]) AND (NOT "ROLL_State".M[110, 4]) AND (NOT "ROLL_State".M[110, 5]) AND (NOT "ROLL_State".M[110, 6]) AND "ROLL_State".M[44, 4]) OR ((NOT "ROLL_State".M[110, 4]) AND (NOT "ROLL_State".M[110, 5]) AND (NOT "ROLL_State".M[110, 6]) AND "ROLL_State".M[46, 1]) OR ((NOT "ROLL_State".M[110, 5]) AND (NOT "ROLL_State".M[110, 6]) AND "ROLL_State".M[47, 4]) OR ((NOT "ROLL_State".M[110, 6]) AND "ROLL_State".M[49, 0]) OR "ROLL_State".M[50, 4]);
   "ROLL_State".M[240, 1] := #r;
   // PB10, STEP 5 network 39
   #r := ((NOT "ROLL_IO".Input[120, 1]) AND ("ROLL_State".M[240, 0] OR "ROLL_State".M[240, 1]) AND "ROLL_IO".Input[12, 5] AND "ROLL_IO".Input[12, 7] AND "ROLL_State".M[110, 7] AND "ROLL_State".M[35, 2] AND "ROLL_State".M[63, 1]);
   IF #r THEN
       "ROLL_State".M[50, 6] := TRUE;
   END_IF;
   #r := ("ROLL_State".M[32, 2] OR "ROLL_State".M[50, 7]);
   IF #r THEN
       "ROLL_State".M[50, 6] := FALSE;
   END_IF;
   // PB10, STEP 5 network 40
   #r := ("ROLL_IO".Input[11, 6] AND "ROLL_IO".Input[120, 1] AND "ROLL_State".M[35, 2] AND "ROLL_State".M[50, 6]);
   IF #r THEN
       "ROLL_State".M[50, 7] := TRUE;
   END_IF;
   #r := ("ROLL_State".M[32, 2] OR "ROLL_State".M[51, 0]);
   IF #r THEN
       "ROLL_State".M[50, 7] := FALSE;
   END_IF;
   // PB10, STEP 5 network 41
   #r := ((NOT "ROLL_IO".Input[12, 1]) AND "ROLL_IO".Input[12, 5] AND "ROLL_State".M[35, 2] AND "ROLL_State".M[50, 7]);
   IF #r THEN
       "ROLL_State".M[51, 0] := TRUE;
   END_IF;
   #r := ("ROLL_State".M[32, 2] OR "ROLL_State".M[51, 1]);
   IF #r THEN
       "ROLL_State".M[51, 0] := FALSE;
   END_IF;
   // PB10, STEP 5 network 42
   #r := ("ROLL_State".M[35, 2] AND "ROLL_State".M[51, 0] AND "ROLL_State".M[80, 6]);
   IF #r THEN
       "ROLL_State".M[51, 1] := TRUE;
   END_IF;
   #r := ("ROLL_State".M[32, 2] OR "ROLL_State".M[51, 2]);
   IF #r THEN
       "ROLL_State".M[51, 1] := FALSE;
   END_IF;
   // PB10, STEP 5 network 43
   #r := ("ROLL_State".M[35, 2] AND "ROLL_State".M[51, 1] AND "ROLL_State".S5Timers[1].Q);
   IF #r THEN
       "ROLL_State".M[51, 2] := TRUE;
   END_IF;
   #r := ("ROLL_State".M[32, 2] OR "ROLL_State".M[51, 3]);
   IF #r THEN
       "ROLL_State".M[51, 2] := FALSE;
   END_IF;
   // PB10, STEP 5 network 44
   #r := ((NOT "ROLL_IO".Input[12, 5]) AND "ROLL_State".M[35, 2] AND "ROLL_State".M[51, 2]);
   IF #r THEN
       "ROLL_State".M[51, 3] := TRUE;
   END_IF;
   #r := ("ROLL_State".M[32, 2] OR "ROLL_State".M[51, 4]);
   IF #r THEN
       "ROLL_State".M[51, 3] := FALSE;
   END_IF;
   // PB10, STEP 5 network 45
   #r := ("ROLL_IO".Input[12, 5] AND "ROLL_IO".Input[12, 7] AND "ROLL_State".M[35, 2] AND "ROLL_State".M[51, 3]);
   IF #r THEN
       "ROLL_State".M[51, 4] := TRUE;
   END_IF;
   #r := ("ROLL_State".M[32, 2] OR "ROLL_State".M[51, 5]);
   IF #r THEN
       "ROLL_State".M[51, 4] := FALSE;
   END_IF;
   // PB10, STEP 5 network 46
   #r := ("ROLL_State".M[35, 2] AND "ROLL_State".M[51, 4]);
   IF #r THEN
       "ROLL_State".M[51, 5] := TRUE;
   END_IF;
   #r := ("ROLL_State".M[32, 2] OR "ROLL_State".M[51, 6]);
   IF #r THEN
       "ROLL_State".M[51, 5] := FALSE;
   END_IF;
   // PB10, STEP 5 network 47
   #r := ("ROLL_IO".Input[13, 3] AND "ROLL_State".M[35, 2] AND "ROLL_State".M[51, 5] AND "ROLL_State".M[63, 1]);
   IF #r THEN
       "ROLL_State".M[51, 6] := TRUE;
   END_IF;
   #r := ("ROLL_State".M[32, 2] OR "ROLL_State".M[52, 0]);
   IF #r THEN
       "ROLL_State".M[51, 6] := FALSE;
   END_IF;
   // PB10, STEP 5 network 48
   #r := (((NOT "ROLL_State".M[110, 1]) AND (NOT "ROLL_State".M[110, 2]) AND (NOT "ROLL_State".M[110, 3]) AND (NOT "ROLL_State".M[110, 4]) AND (NOT "ROLL_State".M[110, 5]) AND (NOT "ROLL_State".M[110, 6]) AND (NOT "ROLL_State".M[110, 7]) AND "ROLL_State".M[41, 4]) OR ((NOT "ROLL_State".M[110, 2]) AND (NOT "ROLL_State".M[110, 3]) AND (NOT "ROLL_State".M[110, 4]) AND (NOT "ROLL_State".M[110, 5]) AND (NOT "ROLL_State".M[110, 6]) AND (NOT "ROLL_State".M[110, 7]) AND "ROLL_State".M[43, 0]));
   "ROLL_State".M[240, 0] := #r;
   // PB10, STEP 5 network 49
   #r := (((NOT "ROLL_State".M[110, 3]) AND (NOT "ROLL_State".M[110, 4]) AND (NOT "ROLL_State".M[110, 5]) AND (NOT "ROLL_State".M[110, 6]) AND (NOT "ROLL_State".M[110, 7]) AND "ROLL_State".M[44, 4]) OR ((NOT "ROLL_State".M[110, 4]) AND (NOT "ROLL_State".M[110, 5]) AND (NOT "ROLL_State".M[110, 6]) AND (NOT "ROLL_State".M[110, 7]) AND "ROLL_State".M[46, 1]) OR ((NOT "ROLL_State".M[110, 5]) AND (NOT "ROLL_State".M[110, 6]) AND (NOT "ROLL_State".M[110, 7]) AND "ROLL_State".M[47, 4]) OR ((NOT "ROLL_State".M[110, 6]) AND (NOT "ROLL_State".M[110, 7]) AND "ROLL_State".M[49, 0]) OR ((NOT "ROLL_State".M[110, 7]) AND "ROLL_State".M[50, 4]) OR "ROLL_State".M[51, 6]);
   "ROLL_State".M[240, 1] := #r;
   // PB10, STEP 5 network 50
   #r := ((NOT "ROLL_IO".Input[11, 0]) AND ("ROLL_State".M[240, 0] OR "ROLL_State".M[240, 1]) AND "ROLL_IO".Input[12, 5] AND "ROLL_IO".Input[12, 7] AND "ROLL_IO".Input[13, 3] AND "ROLL_State".M[35, 2] AND "ROLL_State".M[63, 1]);
   IF #r THEN
       "ROLL_State".M[52, 0] := TRUE;
   END_IF;
   #r := ("ROLL_State".M[32, 2] OR "ROLL_State".M[52, 1]);
   IF #r THEN
       "ROLL_State".M[52, 0] := FALSE;
   END_IF;
   // PB10, STEP 5 network 51
   #r := ("ROLL_IO".Input[11, 0] AND "ROLL_IO".Input[11, 6] AND "ROLL_State".M[35, 2] AND "ROLL_State".M[52, 0]);
   IF #r THEN
       "ROLL_State".M[52, 1] := TRUE;
   END_IF;
   #r := ("ROLL_State".M[32, 2] OR "ROLL_State".M[52, 2]);
   IF #r THEN
       "ROLL_State".M[52, 1] := FALSE;
   END_IF;
   // PB10, STEP 5 network 52
   #r := ((NOT "ROLL_IO".Input[12, 1]) AND (("ROLL_IO".Input[124, 2] AND "ROLL_IO".Input[124, 5]) OR "ROLL_State".M[0, 4]) AND "ROLL_IO".Input[12, 5] AND "ROLL_State".M[35, 2] AND "ROLL_State".M[52, 1]);
   IF #r THEN
       "ROLL_State".M[52, 2] := TRUE;
   END_IF;
   #r := ("ROLL_State".M[32, 2] OR "ROLL_State".M[52, 3]);
   IF #r THEN
       "ROLL_State".M[52, 2] := FALSE;
   END_IF;
   // PB10, STEP 5 network 53
   #r := ("ROLL_IO".Input[12, 1] AND "ROLL_IO".Input[12, 7] AND "ROLL_State".M[35, 2] AND "ROLL_State".M[52, 2]);
   IF #r THEN
       "ROLL_State".M[52, 3] := TRUE;
   END_IF;
   #r := ("ROLL_State".M[32, 2] OR "ROLL_State".M[53, 0] OR "ROLL_State".M[53, 6]);
   IF #r THEN
       "ROLL_State".M[52, 3] := FALSE;
   END_IF;
   // PB10, STEP 5 network 54
   #r := ((NOT "ROLL_IO".Output[113, 3]) AND (NOT "ROLL_IO".Input[123, 5]) AND (NOT "ROLL_IO".Input[123, 6]) AND (NOT "ROLL_IO".Input[124, 1]) AND (NOT "ROLL_State".M[70, 3]) AND "ROLL_IO".Output[113, 2] AND "ROLL_IO".Input[124, 2] AND "ROLL_State".M[0, 3] AND "ROLL_State".M[35, 2] AND "ROLL_State".M[52, 3]);
   IF #r THEN
       "ROLL_State".M[53, 0] := TRUE;
   END_IF;
   #r := ("ROLL_State".M[32, 2] OR "ROLL_State".M[53, 1]);
   IF #r THEN
       "ROLL_State".M[53, 0] := FALSE;
   END_IF;
   // PB10, STEP 5 network 55
   #r := ((NOT "ROLL_IO".Input[124, 2]) AND "ROLL_IO".Input[124, 1] AND "ROLL_State".M[35, 2] AND "ROLL_State".M[53, 0]);
   IF #r THEN
       "ROLL_State".M[53, 1] := TRUE;
   END_IF;
   #r := ("ROLL_State".M[32, 2] OR "ROLL_State".M[53, 2]);
   IF #r THEN
       "ROLL_State".M[53, 1] := FALSE;
   END_IF;
   // PB10, STEP 5 network 56
   #r := ((NOT "ROLL_IO".Input[124, 4]) AND "ROLL_IO".Input[124, 5] AND "ROLL_State".M[35, 2] AND "ROLL_State".M[53, 1]);
   IF #r THEN
       "ROLL_State".M[53, 2] := TRUE;
   END_IF;
   #r := ("ROLL_State".M[32, 2] OR "ROLL_State".M[53, 3]);
   IF #r THEN
       "ROLL_State".M[53, 2] := FALSE;
   END_IF;
   // PB10, STEP 5 network 57
   #r := ((NOT "ROLL_IO".Input[124, 5]) AND "ROLL_IO".Input[124, 4] AND "ROLL_State".M[35, 2] AND "ROLL_State".M[53, 2]);
   IF #r THEN
       "ROLL_State".M[53, 3] := TRUE;
   END_IF;
   #r := ("ROLL_State".M[32, 2] OR "ROLL_State".M[53, 4]);
   IF #r THEN
       "ROLL_State".M[53, 3] := FALSE;
   END_IF;
   // PB10, STEP 5 network 58
   #r := ((NOT "ROLL_State".M[53, 2]) AND "ROLL_State".M[35, 2] AND "ROLL_State".M[53, 3]);
   IF #r THEN
       "ROLL_State".M[53, 4] := TRUE;
   END_IF;
   #r := ("ROLL_State".M[32, 2] OR "ROLL_State".M[53, 5]);
   IF #r THEN
       "ROLL_State".M[53, 4] := FALSE;
   END_IF;
   // PB10, STEP 5 network 59
   #r := ((NOT "ROLL_IO".Input[123, 5]) AND (NOT "ROLL_IO".Input[123, 6]) AND (NOT "ROLL_State".M[70, 3]) AND "ROLL_State".M[35, 2] AND "ROLL_State".M[53, 4]);
   IF #r THEN
       "ROLL_State".M[53, 5] := TRUE;
   END_IF;
   #r := ("ROLL_State".M[32, 2] OR "ROLL_State".M[53, 6]);
   IF #r THEN
       "ROLL_State".M[53, 5] := FALSE;
   END_IF;
   // PB10, STEP 5 network 60
   #r := (("ROLL_State".M[52, 3] OR "ROLL_State".M[53, 5]) AND "ROLL_State".M[35, 2]);
   IF #r THEN
       "ROLL_State".M[53, 6] := TRUE;
   END_IF;
   #r := ("ROLL_State".M[32, 2] OR "ROLL_State".M[37, 0]);
   IF #r THEN
       "ROLL_State".M[53, 6] := FALSE;
   END_IF;
   // PB10, STEP 5 network 61
   RETURN;
END_FUNCTION

FUNCTION "ROLL_PB13" : Void   // FC21, SCL
{ S7_Optimized_Access := 'TRUE' }
VERSION : 0.1
// stored: AutoNumber true, IsIECCheckEnabled false, SetENOAutomatically false, UDAEnableTagReadback false
   VAR_TEMP
      r : Bool;
      a1 : Word;
      a2 : Word;
      activeDataBlock : Int;
      comparisonResults : Array[0..0] of Bool;
   END_VAR
BEGIN

   #r := FALSE;
   #a1 := W#16#0000;
   #a2 := W#16#0000;
   #activeDataBlock := 0;
   // PB13, STEP 5 network 1
   #r := ((NOT "ROLL_State".M[58, 6]) AND ("ROLL_IO".Input[11, 1] OR "ROLL_IO".Input[11, 2] OR "ROLL_IO".Input[11, 3] OR "ROLL_IO".Input[11, 4] OR "ROLL_IO".Input[119, 6] OR "ROLL_IO".Input[119, 7] OR "ROLL_IO".Input[120, 0]) AND "ROLL_IO".Input[11, 6]);
   IF #r THEN
       "ROLL_State".M[58, 7] := TRUE;
   END_IF;
   #r := (((NOT "ROLL_IO".Input[11, 6]) AND ("ROLL_IO".Input[11, 1] OR "ROLL_IO".Input[11, 2] OR "ROLL_IO".Input[11, 3] OR "ROLL_IO".Input[11, 4] OR "ROLL_IO".Input[119, 6] OR "ROLL_IO".Input[119, 7] OR "ROLL_IO".Input[120, 0]) AND "ROLL_IO".Output[23, 0] AND "ROLL_State".M[58, 6]) OR "ROLL_IO".Input[11, 0]);
   IF #r THEN
       "ROLL_State".M[58, 7] := FALSE;
   END_IF;
   // PB13, STEP 5 network 2
   #r := "ROLL_IO".Input[11, 6];
   "ROLL_State".M[58, 6] := #r;
   // PB13, STEP 5 network 3
   #r := (((((NOT "ROLL_IO".Input[11, 0]) OR "ROLL_State".M[80, 7]) AND "ROLL_IO".Input[11, 6]) OR "ROLL_State".M[58, 7]) AND "ROLL_IO".Input[14, 0]);
   "ROLL_State".M[60, 0] := #r;
   // PB13, STEP 5 network 4
   #a2 := #a1;
   #a1 := W#16#2030;
   #r := ((NOT "ROLL_IO".Input[13, 3]) AND "ROLL_IO".Output[24, 0]);
   "ROLL_TimerOp"(Number := 110,
                  Operation := 0,
                  Signal := #r,
                  Preset := #a1);
   // PB13, STEP 5 network 5
   #r := (((NOT "ROLL_State".M[111, 1]) AND (NOT "ROLL_State".M[111, 2]) AND (NOT "ROLL_State".M[111, 5]) AND "ROLL_IO".Input[0, 2] AND "ROLL_State".M[111, 0]) OR ((NOT "ROLL_State".M[61, 5]) AND "ROLL_IO".Input[0, 1] AND "ROLL_State".M[23, 2]) OR ("ROLL_IO".Input[12, 1] AND "ROLL_State".M[111, 5]));
   "ROLL_State".M[60, 1] := #r;
   // PB13, STEP 5 network 6
   #r := (((NOT "ROLL_IO".Input[12, 1]) AND "ROLL_State".M[111, 5]) OR ((NOT "ROLL_State".M[111, 0]) AND (NOT "ROLL_State".M[111, 2]) AND (NOT "ROLL_State".M[111, 5]) AND "ROLL_IO".Input[0, 2] AND "ROLL_State".M[111, 1]) OR ("ROLL_IO".Input[0, 1] AND "ROLL_State".M[23, 3]));
   "ROLL_State".M[60, 3] := #r;
   // PB13, STEP 5 network 7
   #r := (((NOT "ROLL_State".M[111, 0]) AND (NOT "ROLL_State".M[111, 1]) AND (NOT "ROLL_State".M[111, 5]) AND "ROLL_IO".Input[0, 2] AND "ROLL_State".M[111, 2]) OR ((NOT "ROLL_State".M[61, 5]) AND "ROLL_IO".Input[0, 1] AND "ROLL_State".M[0, 3]));
   "ROLL_State".M[60, 2] := #r;
   // PB13, STEP 5 network 8
   #a2 := #a1;
   #a1 := W#16#0005;
   #r := (NOT "ROLL_State".S5Timers[114].Q);
   "ROLL_TimerOp"(Number := 113,
                  Operation := 0,
                  Signal := #r,
                  Preset := #a1);
   #a2 := #a1;
   #a1 := W#16#0005;
   #r := "ROLL_State".S5Timers[113].Q;
   "ROLL_TimerOp"(Number := 114,
                  Operation := 1,
                  Signal := #r,
                  Preset := #a1);
   // PB13, STEP 5 network 9
   #activeDataBlock := 15;
   // PB13, STEP 5 network 10
   #a2 := #a1;
   #a1 := "ROLL_GetDW"(DbNumber := #activeDataBlock, Index := 116);
   #r := ((NOT "ROLL_State".S5Timers[117].Q) AND "ROLL_State".M[62, 4]);
   "ROLL_TimerOp"(Number := 116,
                  Operation := 0,
                  Signal := #r,
                  Preset := #a1);
   #a2 := #a1;
   #a1 := "ROLL_GetDW"(DbNumber := #activeDataBlock, Index := 117);
   #r := "ROLL_State".S5Timers[116].Q;
   "ROLL_TimerOp"(Number := 117,
                  Operation := 1,
                  Signal := #r,
                  Preset := #a1);
   // PB13, STEP 5 network 11
   #activeDataBlock := 19;
   // PB13, STEP 5 network 12
   #r := ("ROLL_IO".Output[24, 2] AND "ROLL_State".M[60, 4] AND "ROLL_State".S5Timers[114].Q);
   "ROLL_CounterOp"(Number := 1,
                    Operation := 3,
                    Signal := #r,
                    Preset := #a1);
   #a2 := #a1;
   #a1 := "ROLL_GetDW"(DbNumber := #activeDataBlock, Index := 1);
   #r := ((((NOT "ROLL_IO".Input[13, 3]) AND (NOT ("ROLL_State".S5Counters[1].Value <> 0)) AND (NOT ("ROLL_State".S5Counters[2].Value <> 0))) OR "ROLL_IO".Input[13, 3] OR "ROLL_State".M[60, 5]) AND "ROLL_State".S5Timers[114].Q);
   "ROLL_CounterOp"(Number := 1,
                    Operation := 0,
                    Signal := #r,
                    Preset := #a1);
   // PB13, STEP 5 network 13
   #r := ("ROLL_IO".Output[24, 0] AND "ROLL_State".M[60, 5] AND "ROLL_State".S5Timers[114].Q);
   "ROLL_CounterOp"(Number := 2,
                    Operation := 3,
                    Signal := #r,
                    Preset := #a1);
   #a2 := #a1;
   #a1 := "ROLL_GetDW"(DbNumber := #activeDataBlock, Index := 2);
   #r := (("ROLL_IO".Input[13, 3] OR "ROLL_State".M[60, 4]) AND "ROLL_State".S5Timers[114].Q);
   "ROLL_CounterOp"(Number := 2,
                    Operation := 0,
                    Signal := #r,
                    Preset := #a1);
   // PB13, STEP 5 network 14
   #r := ((NOT "ROLL_IO".Input[13, 3]) AND "ROLL_IO".Output[24, 2] AND "ROLL_State".M[60, 6]);
   IF #r THEN
       "ROLL_State".M[60, 4] := TRUE;
   END_IF;
   #r := "ROLL_IO".Input[13, 3];
   IF #r THEN
       "ROLL_State".M[60, 4] := FALSE;
   END_IF;
   // PB13, STEP 5 network 15
   #r := ((NOT "ROLL_IO".Input[13, 3]) AND "ROLL_IO".Output[24, 0] AND "ROLL_State".M[60, 6]);
   IF #r THEN
       "ROLL_State".M[60, 5] := TRUE;
   END_IF;
   #r := "ROLL_IO".Input[13, 3];
   IF #r THEN
       "ROLL_State".M[60, 5] := FALSE;
   END_IF;
   // PB13, STEP 5 network 16
   #r := "ROLL_IO".Input[13, 3];
   IF #r THEN
       "ROLL_State".M[60, 6] := TRUE;
   END_IF;
   #r := ("ROLL_State".M[60, 4] OR "ROLL_State".M[60, 5]);
   IF #r THEN
       "ROLL_State".M[60, 6] := FALSE;
   END_IF;
   // PB13, STEP 5 network 17
   #r := ((NOT ("ROLL_State".S5Counters[2].Value <> 0)) AND "ROLL_State".M[62, 6]);
   IF #r THEN
       "ROLL_State".M[60, 7] := TRUE;
   END_IF;
   #r := (NOT "ROLL_State".M[62, 6]);
   IF #r THEN
       "ROLL_State".M[60, 7] := FALSE;
   END_IF;
   // PB13, STEP 5 network 18
   #r := ((NOT "ROLL_IO".Input[13, 3]) AND (NOT ("ROLL_State".S5Counters[1].Value <> 0)) AND "ROLL_State".M[61, 1]);
   IF #r THEN
       "ROLL_State".M[61, 0] := TRUE;
   END_IF;
   #r := (NOT "ROLL_State".M[62, 6]);
   IF #r THEN
       "ROLL_State".M[61, 0] := FALSE;
   END_IF;
   // PB13, STEP 5 network 19
   #r := ("ROLL_State".S5Counters[1].Value <> 0);
   "ROLL_State".M[61, 1] := #r;
   // PB13, STEP 5 network 20
   #r := (("ROLL_State".M[60, 7] OR "ROLL_State".M[62, 6]) AND "ROLL_State".M[61, 0]);
   "ROLL_State".M[61, 2] := #r;
   // PB13, STEP 5 network 21
   #r := ((NOT "ROLL_State".M[61, 6]) AND "ROLL_State".M[60, 1] AND "ROLL_State".M[61, 7]);
   IF #r THEN
       "ROLL_State".M[61, 3] := TRUE;
   END_IF;
   #r := (NOT "ROLL_State".M[61, 7]);
   IF #r THEN
       "ROLL_State".M[61, 3] := FALSE;
   END_IF;
   // PB13, STEP 5 network 22
   #r := ((NOT "ROLL_State".M[61, 6]) AND "ROLL_State".M[60, 2] AND "ROLL_State".M[61, 7]);
   IF #r THEN
       "ROLL_State".M[61, 4] := TRUE;
   END_IF;
   #r := (NOT "ROLL_State".M[61, 7]);
   IF #r THEN
       "ROLL_State".M[61, 4] := FALSE;
   END_IF;
   // PB13, STEP 5 network 23
   #r := ((NOT "ROLL_State".M[61, 6]) AND "ROLL_State".M[60, 3] AND "ROLL_State".M[61, 7]);
   IF #r THEN
       "ROLL_State".M[61, 5] := TRUE;
   END_IF;
   #r := (NOT "ROLL_State".M[61, 7]);
   IF #r THEN
       "ROLL_State".M[61, 5] := FALSE;
   END_IF;
   // PB13, STEP 5 network 24
   #r := "ROLL_State".M[61, 7];
   "ROLL_State".M[61, 6] := #r;
   // PB13, STEP 5 network 25
   #r := (((NOT "ROLL_State".M[111, 5]) AND "ROLL_State".M[37, 3]) OR ((((NOT "ROLL_IO".Input[12, 1]) AND ("ROLL_State".M[41, 0] OR "ROLL_State".M[42, 4] OR "ROLL_State".M[44, 0])) OR (("ROLL_State".M[40, 5] OR "ROLL_State".M[42, 1] OR "ROLL_State".M[43, 5]) AND "ROLL_IO".Input[12, 1])) AND "ROLL_State".M[111, 5]));
   IF #r THEN
       "ROLL_State".M[61, 7] := TRUE;
   END_IF;
   #r := (((NOT "ROLL_IO".Input[12, 5]) AND "ROLL_IO".Input[11, 0] AND "ROLL_State".M[190, 5] AND "ROLL_State".M[20, 1]) OR (("ROLL_State".M[42, 0] OR "ROLL_State".M[43, 4] OR "ROLL_State".M[58, 5]) AND "ROLL_State".M[111, 5]) OR "ROLL_State".M[53, 6]);
   IF #r THEN
       "ROLL_State".M[61, 7] := FALSE;
   END_IF;
   // PB13, STEP 5 network 26
   #r := ((NOT "ROLL_IO".Input[11, 0]) AND (((NOT "ROLL_IO".Input[12, 1]) AND "ROLL_IO".Output[23, 5]) OR ("ROLL_IO".Output[23, 4] AND "ROLL_IO".Input[12, 1])) AND ("ROLL_State".M[61, 3] OR "ROLL_State".M[61, 4] OR "ROLL_State".M[61, 5]));
   IF #r THEN
       "ROLL_State".M[62, 0] := TRUE;
   END_IF;
   #r := ((("ROLL_State".M[41, 3] OR "ROLL_State".M[42, 7] OR "ROLL_State".M[44, 3] OR "ROLL_State".M[46, 0] OR "ROLL_State".M[47, 3] OR "ROLL_State".M[48, 7] OR "ROLL_State".M[50, 3] OR "ROLL_State".M[51, 5]) AND "ROLL_IO".Input[13, 3] AND "ROLL_State".S5Timers[114].Q) OR (NOT "ROLL_State".M[31, 5]) OR (NOT "ROLL_State".M[61, 7]));
   IF #r THEN
       "ROLL_State".M[62, 0] := FALSE;
   END_IF;
   // PB13, STEP 5 network 27
   #r := (((NOT "ROLL_IO".Input[11, 0]) AND ((("ROLL_IO".Input[11, 1] OR "ROLL_IO".Input[11, 2] OR "ROLL_IO".Input[11, 3] OR "ROLL_IO".Input[11, 4] OR "ROLL_IO".Input[119, 6] OR "ROLL_IO".Input[119, 7] OR "ROLL_IO".Input[120, 0]) AND ("ROLL_State".M[80, 6] OR "ROLL_State".M[80, 7])) OR ("ROLL_State".M[60, 0] AND "ROLL_State".M[80, 7]))) OR ("ROLL_IO".Input[11, 0] AND "ROLL_IO".Input[11, 6] AND "ROLL_State".M[80, 7]));
   "ROLL_State".M[62, 1] := #r;
   // PB13, STEP 5 network 28
   #r := (("ROLL_State".M[0, 3] AND "ROLL_State".M[45, 6]) OR "ROLL_State".M[41, 1] OR "ROLL_State".M[42, 5] OR "ROLL_State".M[44, 1] OR "ROLL_State".M[47, 1] OR "ROLL_State".M[48, 5] OR "ROLL_State".M[50, 1]);
   "ROLL_State".M[63, 5] := #r;
   // PB13, STEP 5 network 29
   #r := (((((NOT "ROLL_State".M[60, 1]) AND (NOT "ROLL_State".M[60, 2]) AND (NOT "ROLL_State".M[60, 3]) AND (NOT "ROLL_State".M[63, 1]) AND "ROLL_State".M[74, 0]) OR ((NOT "ROLL_State".M[60, 1]) AND (NOT "ROLL_State".M[60, 2]) AND "ROLL_State".M[60, 3])) AND ("ROLL_State".M[20, 1] OR "ROLL_State".M[20, 2] OR "ROLL_State".M[23, 3]) AND "ROLL_IO".Input[0, 1]) OR ((((NOT "ROLL_State".M[61, 3]) AND (NOT "ROLL_State".M[61, 4]) AND (NOT "ROLL_State".M[61, 5]) AND "ROLL_State".M[62, 6]) OR ((NOT "ROLL_State".M[61, 3]) AND (NOT "ROLL_State".M[61, 4]) AND "ROLL_State".M[61, 5])) AND "ROLL_IO".Input[0, 2]));
   "ROLL_State".M[62, 2] := #r;
   // PB13, STEP 5 network 30
   #r := (((NOT "ROLL_State".M[60, 2]) AND (NOT "ROLL_State".M[60, 3]) AND ("ROLL_State".M[20, 1] OR "ROLL_State".M[23, 2]) AND "ROLL_IO".Input[0, 1] AND "ROLL_State".M[60, 1]) OR ((NOT "ROLL_State".M[61, 4]) AND (NOT "ROLL_State".M[61, 5]) AND (NOT "ROLL_State".M[63, 5]) AND "ROLL_IO".Input[0, 2] AND "ROLL_State".M[61, 3]));
   "ROLL_State".M[62, 3] := #r;
   // PB13, STEP 5 network 31
   #r := (((NOT "ROLL_State".M[60, 1]) AND (NOT "ROLL_State".M[60, 3]) AND ("ROLL_State".M[0, 3] OR "ROLL_State".M[20, 1]) AND "ROLL_IO".Input[0, 1] AND "ROLL_State".M[60, 2]) OR ((((NOT "ROLL_State".M[61, 3]) AND (NOT "ROLL_State".M[61, 5]) AND "ROLL_State".M[61, 4]) OR ("ROLL_State".M[61, 3] AND "ROLL_State".M[63, 5])) AND "ROLL_IO".Input[0, 2]));
   "ROLL_State".M[62, 4] := #r;
   // PB13, STEP 5 network 32
   #r := ((((NOT "ROLL_State".M[190, 5]) AND ("ROLL_State".M[0, 3] OR "ROLL_State".M[23, 2] OR "ROLL_State".M[23, 3]) AND ("ROLL_State".M[60, 1] OR "ROLL_State".M[60, 2] OR "ROLL_State".M[60, 3]) AND "ROLL_IO".Input[0, 1] AND "ROLL_State".M[190, 6] AND "ROLL_State".M[62, 1]) OR ("ROLL_IO".Input[0, 2] AND "ROLL_State".M[31, 5] AND "ROLL_State".M[62, 0])) AND ("ROLL_State".M[62, 5] OR "ROLL_State".S5Timers[114].Q) AND "ROLL_State".M[60, 0]);
   "ROLL_State".M[62, 5] := #r;
   // PB13, STEP 5 network 33
   #r := ((NOT "ROLL_State".M[63, 1]) AND (((NOT "ROLL_State".M[62, 0]) AND "ROLL_IO".Input[0, 2] AND "ROLL_State".M[31, 5]) OR ((((NOT "ROLL_State".M[190, 6]) AND ("ROLL_State".M[0, 3] OR "ROLL_State".M[20, 2] OR "ROLL_State".M[23, 2] OR "ROLL_State".M[23, 3]) AND "ROLL_State".M[190, 5]) OR "ROLL_State".M[74, 0]) AND "ROLL_IO".Input[0, 1] AND "ROLL_State".M[62, 1])) AND ("ROLL_State".M[62, 6] OR "ROLL_State".S5Timers[114].Q) AND "ROLL_State".M[60, 0]);
   "ROLL_State".M[62, 6] := #r;
   // PB13, STEP 5 network 34
   #r := ((((NOT "ROLL_State".M[61, 2]) AND (NOT "ROLL_State".M[63, 1]) AND "ROLL_State".M[62, 6]) OR "ROLL_State".M[62, 5]) AND (((NOT "ROLL_State".M[62, 2]) AND (NOT "ROLL_State".M[62, 4]) AND (NOT "ROLL_State".M[62, 6]) AND "ROLL_State".M[62, 3]) OR ((NOT "ROLL_State".M[62, 6]) AND ("ROLL_IO".Input[13, 3] OR "ROLL_State".S5Timers[117].Q) AND "ROLL_State".M[62, 4]) OR (((NOT "ROLL_State".M[62, 4]) OR "ROLL_State".M[62, 6]) AND ("ROLL_State".S5Counters[1].Value <> 0))) AND ("ROLL_State".M[62, 2] OR "ROLL_State".M[62, 3] OR "ROLL_State".M[62, 4]));
   "ROLL_State".M[62, 7] := #r;
   // PB13, STEP 5 network 35
   #r := ((NOT "ROLL_IO".Output[24, 0]) AND (NOT "ROLL_State".M[5, 1]) AND (NOT "ROLL_State".M[63, 4]) AND ((NOT "ROLL_State".S5Timers[115].Q) OR "ROLL_IO".Output[24, 2]) AND "ROLL_IO".Input[13, 5] AND "ROLL_State".M[29, 0] AND "ROLL_State".M[60, 0] AND "ROLL_State".M[62, 7]);
   "ROLL_IO".Output[24, 2] := #r;
   // PB13, STEP 5 network 36
   #r := ((((NOT "ROLL_State".M[62, 2]) AND (NOT "ROLL_State".M[62, 6])) OR ("ROLL_State".S5Counters[2].Value <> 0)) AND (((NOT "ROLL_State".M[63, 1]) AND "ROLL_State".M[62, 6]) OR "ROLL_State".M[62, 5]) AND ((NOT "ROLL_State".M[62, 4]) OR (NOT "ROLL_State".M[62, 5])));
   "ROLL_State".M[63, 0] := #r;
   // PB13, STEP 5 network 37
   #r := ((NOT "ROLL_IO".Output[24, 2]) AND (NOT "ROLL_State".M[5, 1]) AND (NOT "ROLL_State".M[63, 4]) AND ((NOT "ROLL_State".S5Timers[115].Q) OR "ROLL_IO".Output[24, 0]) AND "ROLL_IO".Input[13, 5] AND "ROLL_State".M[29, 0] AND "ROLL_State".M[60, 0] AND "ROLL_State".M[63, 0]);
   "ROLL_IO".Output[24, 0] := #r;
   // PB13, STEP 5 network 38
   #r := ((NOT "ROLL_IO".Output[24, 5]) AND "ROLL_IO".Output[24, 0] AND "ROLL_IO".Input[13, 3]);
   "ROLL_IO".Output[24, 1] := #r;
   // PB13, STEP 5 network 39
   #r := ("ROLL_IO".Output[24, 0] OR "ROLL_IO".Output[24, 2] OR "ROLL_State".M[63, 6]);
   "ROLL_State".M[240, 0] := #r;
   // PB13, STEP 5 network 40
   #r := ((NOT "ROLL_IO".Input[12, 5]) AND (("ROLL_State".M[190, 5] AND "ROLL_State".M[23, 0]) OR "ROLL_State".M[52, 2]) AND "ROLL_IO".Input[11, 0] AND "ROLL_IO".Input[11, 6]);
   IF #r THEN
       "ROLL_State".M[63, 6] := TRUE;
   END_IF;
   #r := (("ROLL_IO".Input[12, 1] OR "ROLL_IO".Input[12, 5]) AND "ROLL_IO".Input[11, 0] AND "ROLL_IO".Input[11, 6] AND "ROLL_IO".Input[12, 7]);
   IF #r THEN
       "ROLL_State".M[63, 6] := FALSE;
   END_IF;
   // PB13, STEP 5 network 41
   #r := ((((NOT "ROLL_State".M[63, 7]) AND "ROLL_IO".Output[24, 0] AND "ROLL_State".S5Timers[111].Q) OR ("ROLL_IO".Input[11, 0] AND "ROLL_State".M[80, 6]) OR (NOT "ROLL_State".S5Timers[11].Q)) AND "ROLL_IO".Input[13, 3]);
   IF #r THEN
       "ROLL_State".M[63, 1] := TRUE;
   END_IF;
   #r := (((NOT "ROLL_IO".Input[13, 3]) AND "ROLL_IO".Input[3, 0] AND "ROLL_State".S5Timers[11].Q) OR "ROLL_IO".Output[24, 2]);
   IF #r THEN
       "ROLL_State".M[63, 1] := FALSE;
   END_IF;
   // PB13, STEP 5 network 42
   #a2 := #a1;
   #a1 := W#16#1030;
   #r := ("ROLL_IO".Output[24, 0] AND "ROLL_IO".Input[13, 3] AND "ROLL_State".M[29, 0] AND "ROLL_State".M[61, 2]);
   "ROLL_TimerOp"(Number := 111,
                  Operation := 0,
                  Signal := #r,
                  Preset := #a1);
   // PB13, STEP 5 network 43
   #r := (((NOT "ROLL_IO".Input[13, 3]) AND "ROLL_IO".Input[0, 1] AND "ROLL_State".M[0, 3] AND "ROLL_State".M[190, 6]) OR ((((NOT "ROLL_State".M[61, 2]) AND "ROLL_State".M[62, 6]) OR "ROLL_State".M[62, 5]) AND ("ROLL_State".M[62, 2] OR "ROLL_State".M[62, 3] OR "ROLL_State".M[62, 4])) OR ("ROLL_IO".Input[13, 3] AND "ROLL_State".M[63, 7]));
   "ROLL_State".M[63, 7] := #r;
   "ROLL_IO".Output[24, 5] := #r;
   // PB13, STEP 5 network 44
   #r := ("ROLL_IO".Output[24, 0] OR "ROLL_IO".Output[24, 2]);
   "ROLL_IO".Output[24, 4] := #r;
   // PB13, STEP 5 network 45
   #r := ("ROLL_State".M[41, 1] OR "ROLL_State".M[42, 5] OR "ROLL_State".M[44, 1] OR "ROLL_State".M[45, 6] OR "ROLL_State".M[47, 1] OR "ROLL_State".M[48, 5] OR "ROLL_State".M[50, 1]);
   "ROLL_State".M[240, 0] := #r;
   // PB13, STEP 5 network 46
   #r := "ROLL_State".M[111, 1];
   "ROLL_State".M[240, 1] := #r;
   // PB13, STEP 5 network 47
   "ROLL_FB69"();
   // PB13, STEP 5 network 48
   #a2 := #a1;
   #a1 := "ROLL_GetM"(FirstByte := 240, Width := 16);
   #r := ("ROLL_IO".Output[24, 0] OR "ROLL_IO".Output[24, 2]);
   "ROLL_TimerOp"(Number := 115,
                  Operation := 1,
                  Signal := #r,
                  Preset := #a1);
   // PB13, STEP 5 network 49
   #r := ((("ROLL_IO".Output[24, 0] AND "ROLL_State".M[60, 5]) OR ("ROLL_IO".Output[24, 2] AND "ROLL_State".M[60, 4])) AND "ROLL_State".S5Timers[114].Q);
   "ROLL_CounterOp"(Number := 3,
                    Operation := 3,
                    Signal := #r,
                    Preset := #a1);
   #r := ((((NOT "ROLL_State".M[60, 4]) AND (NOT "ROLL_State".M[60, 5]) AND ("ROLL_IO".Output[24, 0] OR "ROLL_IO".Output[24, 2])) OR ("ROLL_IO".Output[24, 0] AND "ROLL_State".M[60, 4]) OR ("ROLL_IO".Output[24, 2] AND "ROLL_State".M[60, 5])) AND "ROLL_State".S5Timers[114].Q);
   "ROLL_CounterOp"(Number := 3,
                    Operation := 2,
                    Signal := #r,
                    Preset := #a1);
   #a2 := #a1;
   #a1 := W#16#0500;
   #r := (("ROLL_IO".Input[13, 3] AND "ROLL_State".S5Timers[114].Q) OR ("ROLL_State".M[3, 1] AND "ROLL_State".M[63, 2]));
   "ROLL_CounterOp"(Number := 3,
                    Operation := 0,
                    Signal := #r,
                    Preset := #a1);
   // PB13, STEP 5 network 50
   #a2 := #a1;
   #a1 := INT_TO_WORD("ROLL_State".S5Counters[3].Value);
   #a2 := #a1;
   #a1 := W#16#0208;
   #comparisonResults[0] := (WORD_TO_INT(#a2) > WORD_TO_INT(#a1));
   #r := #comparisonResults[0];
   "ROLL_State".M[63, 2] := #r;
   // PB13, STEP 5 network 51
   #a2 := #a1;
   #a1 := W#16#1060;
   #r := ((("ROLL_IO".Output[24, 0] AND "ROLL_State".M[63, 7]) OR "ROLL_IO".Output[24, 2]) AND "ROLL_IO".Input[13, 3]);
   "ROLL_TimerOp"(Number := 112,
                  Operation := 0,
                  Signal := #r,
                  Preset := #a1);
   // PB13, STEP 5 network 52
   #r := ((NOT ("ROLL_State".S5Counters[2].Value <> 0)) AND "ROLL_State".M[61, 2] AND "ROLL_State".M[62, 6] AND ("ROLL_State".S5Counters[1].Value <> 0));
   "ROLL_State".M[63, 3] := #r;
   // PB13, STEP 5 network 53
   #r := (((NOT "ROLL_IO".Input[0, 4]) AND "ROLL_IO".Input[0, 2] AND "ROLL_State".M[63, 4]) OR "ROLL_State".M[11, 0] OR "ROLL_State".M[11, 1] OR "ROLL_State".M[11, 2] OR "ROLL_State".M[11, 3]);
   "ROLL_State".M[63, 4] := #r;
   // PB13, STEP 5 network 54
   RETURN;
END_FUNCTION

FUNCTION "ROLL_PB14" : Void   // FC22, SCL
{ S7_Optimized_Access := 'TRUE' }
VERSION : 0.1
// stored: AutoNumber true, IsIECCheckEnabled false, SetENOAutomatically false, UDAEnableTagReadback false
   VAR_TEMP
      r : Bool;
      a1 : Word;
      a2 : Word;
      activeDataBlock : Int;
      comparisonResults : Array[0..0] of Bool;
   END_VAR
BEGIN

   #r := FALSE;
   #a1 := W#16#0000;
   #a2 := W#16#0000;
   #activeDataBlock := 0;
   // PB14, STEP 5 network 1
   #activeDataBlock := 15;
   // PB14, STEP 5 network 2
   #r := ((NOT "ROLL_State".M[37, 5]) AND (NOT "ROLL_State".M[53, 2]) AND (NOT "ROLL_State".M[53, 3]) AND (((NOT "ROLL_State".S5Timers[21].Q) AND "ROLL_IO".Input[123, 4] AND "ROLL_State".M[31, 4]) OR ("ROLL_State".M[70, 4] AND "ROLL_State".S5Timers[45].Q) OR "ROLL_State".M[37, 7] OR "ROLL_State".M[53, 4] OR "ROLL_State".M[70, 7]) AND ((NOT "ROLL_State".S5Timers[95].Q) OR "ROLL_State".M[53, 4]) AND "ROLL_State".M[31, 5] AND "ROLL_State".M[35, 2]);
   "ROLL_State".M[64, 0] := #r;
   // PB14, STEP 5 network 3
   #r := (((NOT "ROLL_State".M[31, 4]) AND (NOT "ROLL_State".M[31, 5]) AND "ROLL_IO".Input[125, 4]) OR ((((NOT "ROLL_IO".Output[113, 4]) AND "ROLL_IO".Output[113, 5] AND "ROLL_State".M[72, 1]) OR "ROLL_State".M[53, 4]) AND "ROLL_State".M[31, 5] AND "ROLL_State".M[35, 2]));
   "ROLL_State".M[64, 1] := #r;
   // PB14, STEP 5 network 4
   #r := ("ROLL_IO".Input[123, 4] AND "ROLL_State".S5Timers[20].Q);
   IF #r THEN
       "ROLL_State".M[64, 4] := TRUE;
   END_IF;
   #r := (((NOT "ROLL_IO".Output[113, 3]) AND (NOT "ROLL_IO".Input[123, 4])) OR (NOT "ROLL_State".M[31, 5]));
   IF #r THEN
       "ROLL_State".M[64, 4] := FALSE;
   END_IF;
   // PB14, STEP 5 network 5
   #r := "ROLL_State".M[37, 5];
   IF #r THEN
       "ROLL_State".M[64, 5] := TRUE;
   END_IF;
   #r := ((NOT "ROLL_State".M[31, 5]) OR "ROLL_State".M[39, 5]);
   IF #r THEN
       "ROLL_State".M[64, 5] := FALSE;
   END_IF;
   // PB14, STEP 5 network 6
   #r := ((("ROLL_State".M[40, 2] OR "ROLL_State".M[44, 7] OR "ROLL_State".M[50, 6]) AND "ROLL_State".M[63, 1]) OR "ROLL_State".M[41, 6] OR "ROLL_State".M[43, 2] OR "ROLL_State".M[44, 7] OR "ROLL_State".M[46, 2] OR "ROLL_State".M[47, 6] OR "ROLL_State".M[49, 2]);
   "ROLL_State".M[65, 0] := #r;
   // PB14, STEP 5 network 7
   #r := ("ROLL_IO".Input[12, 5] AND "ROLL_IO".Input[12, 7] AND "ROLL_State".M[52, 0] AND "ROLL_State".M[63, 1]);
   "ROLL_State".M[65, 5] := #r;
   // PB14, STEP 5 network 8
   #r := (((NOT "ROLL_IO".Input[11, 0]) AND "ROLL_State".M[52, 0]) OR ((NOT "ROLL_IO".Input[11, 1]) AND "ROLL_State".M[40, 2]) OR ((NOT "ROLL_IO".Input[11, 2]) AND "ROLL_State".M[41, 6]) OR ((NOT "ROLL_IO".Input[11, 3]) AND "ROLL_State".M[43, 2]) OR ((NOT "ROLL_IO".Input[11, 4]) AND "ROLL_State".M[44, 7]) OR ((NOT "ROLL_IO".Input[119, 6]) AND "ROLL_State".M[46, 2]) OR ((NOT "ROLL_IO".Input[119, 7]) AND "ROLL_State".M[47, 6]) OR ((NOT "ROLL_IO".Input[120, 0]) AND "ROLL_State".M[49, 2]) OR ((NOT "ROLL_IO".Input[120, 1]) AND "ROLL_State".M[50, 6]));
   "ROLL_State".M[65, 6] := #r;
   // PB14, STEP 5 network 9
   #r := (("ROLL_IO".Input[11, 0] AND "ROLL_State".M[40, 0]) OR ("ROLL_IO".Input[11, 1] AND "ROLL_State".M[41, 0]) OR ("ROLL_IO".Input[11, 2] AND "ROLL_State".M[42, 4]) OR ("ROLL_IO".Input[11, 3] AND "ROLL_State".M[44, 0]) OR ("ROLL_IO".Input[11, 4] AND "ROLL_State".M[45, 5]) OR ("ROLL_IO".Input[119, 6] AND "ROLL_State".M[47, 0]) OR ("ROLL_IO".Input[119, 7] AND "ROLL_State".M[48, 4]) OR ("ROLL_IO".Input[120, 0] AND "ROLL_State".M[50, 0]) OR ("ROLL_IO".Input[120, 1] AND "ROLL_State".M[51, 3]));
   "ROLL_State".M[66, 2] := #r;
   // PB14, STEP 5 network 10
   #r := (("ROLL_State".M[66, 2] OR "ROLL_State".M[68, 2]) AND "ROLL_IO".Input[11, 6]);
   "ROLL_State".M[66, 4] := #r;
   // PB14, STEP 5 network 11
   #r := (("ROLL_IO".Input[11, 1] AND "ROLL_State".M[40, 4]) OR ("ROLL_IO".Input[11, 2] AND "ROLL_State".M[42, 0]) OR ("ROLL_IO".Input[11, 3] AND "ROLL_State".M[43, 4]) OR ("ROLL_IO".Input[11, 4] AND "ROLL_State".M[45, 1]) OR ("ROLL_IO".Input[119, 6] AND "ROLL_State".M[46, 4]) OR ("ROLL_IO".Input[119, 7] AND "ROLL_State".M[48, 0]) OR ("ROLL_IO".Input[120, 0] AND "ROLL_State".M[49, 4]) OR ("ROLL_IO".Input[120, 1] AND "ROLL_State".M[51, 0]));
   "ROLL_State".M[66, 5] := #r;
   // PB14, STEP 5 network 12
   #r := (((NOT "ROLL_IO".Input[12, 1]) OR (NOT "ROLL_IO".Input[12, 7])) AND "ROLL_IO".Input[11, 0] AND "ROLL_State".M[52, 2]);
   "ROLL_State".M[66, 6] := #r;
   // PB14, STEP 5 network 13
   #r := (("ROLL_State".M[66, 5] OR "ROLL_State".M[66, 6] OR "ROLL_State".M[68, 3]) AND "ROLL_IO".Input[11, 6]);
   "ROLL_State".M[66, 7] := #r;
   // PB14, STEP 5 network 14
   #r := ((NOT "ROLL_IO".Output[113, 3]) AND (NOT "ROLL_State".M[9, 3]) AND "ROLL_IO".Input[124, 5] AND "ROLL_State".M[39, 6]);
   "ROLL_State".M[67, 0] := #r;
   // PB14, STEP 5 network 15
   #r := ((NOT "ROLL_IO".Output[113, 3]) AND (NOT "ROLL_State".M[9, 3]) AND "ROLL_IO".Input[124, 5] AND "ROLL_State".M[53, 0]);
   "ROLL_State".M[67, 1] := #r;
   // PB14, STEP 5 network 16
   #r := ((NOT "ROLL_IO".Input[124, 5]) AND "ROLL_IO".Input[124, 1] AND "ROLL_State".M[39, 4]);
   "ROLL_State".M[67, 5] := #r;
   // PB14, STEP 5 network 17
   #r := ((NOT "ROLL_IO".Input[124, 4]) AND "ROLL_IO".Input[124, 1] AND "ROLL_State".M[53, 2]);
   "ROLL_State".M[67, 6] := #r;
   // PB14, STEP 5 network 18
   #r := ((("ROLL_IO".Input[5, 1] AND "ROLL_State".M[40, 5]) OR ("ROLL_State".M[0, 3] AND "ROLL_State".M[45, 2]) OR "ROLL_State".M[42, 1] OR "ROLL_State".M[43, 5] OR "ROLL_State".M[46, 5] OR "ROLL_State".M[48, 1] OR "ROLL_State".M[49, 5]) AND "ROLL_State".M[111, 3]);
   "ROLL_State".M[68, 0] := #r;
   // PB14, STEP 5 network 19
   #r := ((NOT "ROLL_State".S5Timers[25].Q) AND (("ROLL_IO".Input[12, 1] AND "ROLL_IO".Input[12, 7]) OR "ROLL_State".M[68, 2]) AND ("ROLL_State".M[68, 2] OR "ROLL_State".S5Timers[24].Q) AND "ROLL_State".M[68, 0]);
   "ROLL_State".M[68, 2] := #r;
   // PB14, STEP 5 network 20
   #r := (((NOT "ROLL_IO".Input[12, 1]) OR (NOT "ROLL_IO".Input[12, 7])) AND ("ROLL_State".M[68, 3] OR "ROLL_State".S5Timers[24].Q) AND "ROLL_State".M[68, 0]);
   "ROLL_State".M[68, 3] := #r;
   // PB14, STEP 5 network 21
   #a2 := #a1;
   #a1 := "ROLL_GetDW"(DbNumber := #activeDataBlock, Index := 24);
   #r := ((NOT "ROLL_State".M[68, 2]) AND (NOT "ROLL_State".M[68, 3]));
   "ROLL_TimerOp"(Number := 24,
                  Operation := 0,
                  Signal := #r,
                  Preset := #a1);
   // PB14, STEP 5 network 22
   #a2 := #a1;
   #a1 := "ROLL_GetDW"(DbNumber := #activeDataBlock, Index := 25);
   #r := "ROLL_State".M[68, 2];
   "ROLL_TimerOp"(Number := 25,
                  Operation := 0,
                  Signal := #r,
                  Preset := #a1);
   // PB14, STEP 5 network 23
   RETURN;
END_FUNCTION

FUNCTION "ROLL_PB15" : Void   // FC23, SCL
{ S7_Optimized_Access := 'TRUE' }
VERSION : 0.1
// stored: AutoNumber true, IsIECCheckEnabled false, SetENOAutomatically false, UDAEnableTagReadback false
   VAR_TEMP
      r : Bool;
      a1 : Word;
      a2 : Word;
      activeDataBlock : Int;
      comparisonResults : Array[0..0] of Bool;
   END_VAR
BEGIN

   #r := FALSE;
   #a1 := W#16#0000;
   #a2 := W#16#0000;
   #activeDataBlock := 0;
   // PB15, STEP 5 network 1
   #r := ((NOT "ROLL_IO".Output[113, 2]) AND "ROLL_IO".Output[113, 3] AND "ROLL_IO".Input[123, 4]);
   IF #r THEN
       "ROLL_State".M[70, 2] := TRUE;
   END_IF;
   #r := (((NOT "ROLL_IO".Input[123, 4]) AND "ROLL_IO".Input[123, 5]) OR "ROLL_State".M[73, 7]);
   IF #r THEN
       "ROLL_State".M[70, 2] := FALSE;
   END_IF;
   // PB15, STEP 5 network 2
   #r := ((((NOT "ROLL_State".M[20, 2]) AND "ROLL_IO".Input[123, 6] AND "ROLL_State".M[74, 0]) OR "ROLL_State".M[71, 0]) AND "ROLL_IO".Output[113, 2] AND "ROLL_IO".Input[124, 1] AND "ROLL_IO".Input[124, 4]);
   IF #r THEN
       "ROLL_State".M[70, 3] := TRUE;
   END_IF;
   #r := (((NOT "ROLL_IO".Input[123, 5]) AND (NOT "ROLL_IO".Input[123, 6])) OR "ROLL_State".M[73, 7]);
   IF #r THEN
       "ROLL_State".M[70, 3] := FALSE;
   END_IF;
   // PB15, STEP 5 network 3
   #r := ((NOT "ROLL_State".M[16, 0]) AND (NOT "ROLL_State".M[16, 1]) AND (NOT "ROLL_State".M[16, 4]) AND (NOT "ROLL_State".M[71, 1]) AND "ROLL_IO".Input[123, 1] AND "ROLL_State".M[191, 4] AND "ROLL_State".M[31, 4] AND "ROLL_State".S5Timers[45].Q);
   IF #r THEN
       "ROLL_State".M[70, 4] := TRUE;
   END_IF;
   #r := ((NOT "ROLL_IO".Input[123, 1]) OR "ROLL_State".M[73, 7]);
   IF #r THEN
       "ROLL_State".M[70, 4] := FALSE;
   END_IF;
   // PB15, STEP 5 network 4
   #r := "ROLL_IO".Input[123, 6];
   IF #r THEN
       "ROLL_State".M[70, 5] := TRUE;
   END_IF;
   #r := ("ROLL_IO".Input[125, 0] OR "ROLL_State".M[73, 7]);
   IF #r THEN
       "ROLL_State".M[70, 5] := FALSE;
   END_IF;
   // PB15, STEP 5 network 5
   #r := ((NOT "ROLL_IO".Input[125, 1]) AND "ROLL_IO".Output[113, 4] AND "ROLL_IO".Input[125, 0]);
   IF #r THEN
       "ROLL_State".M[70, 6] := TRUE;
   END_IF;
   #r := (("ROLL_IO".Output[113, 5] AND "ROLL_IO".Input[125, 1]) OR "ROLL_State".M[73, 7]);
   IF #r THEN
       "ROLL_State".M[70, 6] := FALSE;
   END_IF;
   // PB15, STEP 5 network 6
   #r := ((NOT "ROLL_State".M[71, 1]) AND "ROLL_IO".Input[123, 1] AND "ROLL_State".S5Timers[45].Q);
   IF #r THEN
       "ROLL_State".M[70, 7] := TRUE;
   END_IF;
   #r := ("ROLL_IO".Input[123, 4] OR "ROLL_State".M[73, 7]);
   IF #r THEN
       "ROLL_State".M[70, 7] := FALSE;
   END_IF;
   // PB15, STEP 5 network 7
   #r := ("ROLL_IO".Output[113, 3] AND "ROLL_IO".Input[123, 5]);
   IF #r THEN
       "ROLL_State".M[71, 0] := TRUE;
   END_IF;
   #r := ("ROLL_State".M[70, 3] OR "ROLL_State".M[73, 7]);
   IF #r THEN
       "ROLL_State".M[71, 0] := FALSE;
   END_IF;
   // PB15, STEP 5 network 8
   #r := ((NOT "ROLL_State".M[190, 6]) AND (NOT "ROLL_State".M[28, 4]) AND ("ROLL_State".M[20, 1] OR "ROLL_State".M[20, 2]) AND "ROLL_IO".Input[0, 1] AND "ROLL_State".M[190, 5]);
   "ROLL_State".M[74, 0] := #r;
   // PB15, STEP 5 network 9
   RETURN;
END_FUNCTION

FUNCTION "ROLL_PB16" : Void   // FC24, SCL
{ S7_Optimized_Access := 'TRUE' }
VERSION : 0.1
// stored: AutoNumber true, IsIECCheckEnabled false, SetENOAutomatically false, UDAEnableTagReadback false
   VAR_TEMP
      r : Bool;
      a1 : Word;
      a2 : Word;
      activeDataBlock : Int;
      comparisonResults : Array[0..0] of Bool;
   END_VAR
BEGIN

   #r := FALSE;
   #a1 := W#16#0000;
   #a2 := W#16#0000;
   #activeDataBlock := 0;
   // PB16, STEP 5 network 1
   #r := ("ROLL_IO".Input[0, 1] AND "ROLL_State".M[190, 5] AND "ROLL_State".M[190, 6] AND "ROLL_State".M[27, 7]);
   "ROLL_State".M[73, 7] := #r;
   // PB16, STEP 5 network 2
   #r := (("ROLL_State".M[20, 3] OR "ROLL_State".M[20, 5]) AND "ROLL_IO".Input[124, 1] AND "ROLL_IO".Input[124, 4]);
   "ROLL_State".M[74, 2] := #r;
   // PB16, STEP 5 network 3
   #r := (((NOT "ROLL_State".M[190, 5]) AND "ROLL_State".M[190, 6] AND "ROLL_State".M[74, 2]) OR (("ROLL_State".M[70, 2] OR "ROLL_State".M[70, 3]) AND "ROLL_State".M[74, 0]));
   "ROLL_State".M[74, 1] := #r;
   // PB16, STEP 5 network 4
   #r := (("ROLL_State".M[20, 4] OR "ROLL_State".M[20, 5]) AND "ROLL_IO".Input[0, 1] AND "ROLL_State".M[190, 6]);
   "ROLL_State".M[74, 4] := #r;
   // PB16, STEP 5 network 5
   #r := ((NOT "ROLL_IO".Output[113, 3]) AND ("ROLL_IO".Input[123, 6] OR "ROLL_State".M[70, 3] OR "ROLL_State".M[70, 5] OR "ROLL_State".M[70, 6]) AND ("ROLL_State".M[74, 0] OR "ROLL_State".M[74, 4]));
   "ROLL_State".M[74, 5] := #r;
   // PB16, STEP 5 network 6
   #r := ((NOT "ROLL_IO".Input[11, 0]) AND (NOT "ROLL_IO".Input[11, 1]) AND (NOT "ROLL_IO".Input[11, 2]) AND (NOT "ROLL_IO".Input[11, 3]) AND (NOT "ROLL_IO".Input[11, 4]) AND (NOT "ROLL_IO".Input[119, 6]) AND (NOT "ROLL_IO".Input[119, 7]) AND (NOT "ROLL_IO".Input[120, 0]) AND (NOT "ROLL_IO".Input[120, 1]));
   "ROLL_State".M[75, 2] := #r;
   // PB16, STEP 5 network 7
   #r := (("ROLL_State".M[190, 6] AND "ROLL_State".M[23, 1] AND "ROLL_State".M[75, 3]) OR "ROLL_State".M[75, 2]);
   "ROLL_State".M[75, 3] := #r;
   // PB16, STEP 5 network 8
   #r := ((((NOT "ROLL_IO".Input[11, 0]) AND (NOT "ROLL_IO".Input[11, 1]) AND (NOT "ROLL_IO".Input[11, 2]) AND (NOT "ROLL_IO".Input[11, 3]) AND (NOT "ROLL_IO".Input[11, 4]) AND (NOT "ROLL_IO".Input[119, 6]) AND (NOT "ROLL_IO".Input[119, 7]) AND (NOT "ROLL_IO".Input[120, 0]) AND (NOT "ROLL_IO".Input[120, 1]) AND "ROLL_IO".Input[13, 3]) OR "ROLL_State".M[63, 1]) AND ((NOT "ROLL_IO".Input[11, 6]) OR (NOT "ROLL_State".M[75, 3]) OR "ROLL_State".M[75, 2]) AND "ROLL_IO".Input[0, 1] AND "ROLL_IO".Input[12, 5] AND "ROLL_State".M[190, 6] AND "ROLL_State".M[23, 1]);
   "ROLL_State".M[75, 4] := #r;
   // PB16, STEP 5 network 9
   #r := ((((NOT "ROLL_IO".Input[11, 0]) AND (NOT "ROLL_IO".Input[11, 1]) AND (NOT "ROLL_IO".Input[11, 2]) AND (NOT "ROLL_IO".Input[11, 3]) AND (NOT "ROLL_IO".Input[11, 4]) AND (NOT "ROLL_IO".Input[119, 6]) AND (NOT "ROLL_IO".Input[119, 7]) AND (NOT "ROLL_IO".Input[120, 0]) AND (NOT "ROLL_IO".Input[120, 1]) AND "ROLL_IO".Input[13, 3]) OR "ROLL_State".M[63, 1]) AND (((NOT "ROLL_State".M[190, 6]) AND "ROLL_State".M[190, 5] AND "ROLL_State".M[23, 1]) OR "ROLL_State".M[74, 0]) AND "ROLL_IO".Input[0, 1]);
   "ROLL_State".M[75, 5] := #r;
   // PB16, STEP 5 network 10
   #r := (((NOT "ROLL_IO".Input[11, 0]) AND (("ROLL_IO".Input[0, 1] AND "ROLL_State".M[190, 5] AND "ROLL_State".M[23, 1]) OR "ROLL_State".M[74, 0]) AND "ROLL_State".M[63, 1]) OR ("ROLL_IO".Input[0, 1] AND "ROLL_State".M[190, 6] AND "ROLL_State".M[23, 1] AND "ROLL_State".M[75, 2]));
   "ROLL_State".M[75, 6] := #r;
   // PB16, STEP 5 network 11
   #r := ((NOT "ROLL_IO".Input[11, 0]) AND "ROLL_IO".Input[11, 6] AND "ROLL_State".M[190, 5] AND "ROLL_State".M[23, 0]);
   "ROLL_State".M[76, 0] := #r;
   // PB16, STEP 5 network 12
   #r := (((NOT "ROLL_IO".Input[11, 0]) AND "ROLL_State".M[74, 0]) OR ("ROLL_IO".Input[11, 0] AND "ROLL_IO".Input[11, 6] AND "ROLL_State".M[190, 6] AND "ROLL_State".M[23, 0]));
   "ROLL_State".M[76, 1] := #r;
   // PB16, STEP 5 network 13
   #r := (("ROLL_State".M[76, 0] OR "ROLL_State".M[76, 1]) AND "ROLL_IO".Input[0, 1]);
   "ROLL_State".M[76, 2] := #r;
   // PB16, STEP 5 network 14
   #r := ((NOT "ROLL_IO".Input[12, 1]) AND (NOT "ROLL_IO".Input[12, 5]));
   "ROLL_State".M[240, 0] := #r;
   // PB16, STEP 5 network 15
   #r := (("ROLL_State".M[190, 6] AND "ROLL_State".M[23, 0] AND "ROLL_State".M[77, 1]) OR "ROLL_State".M[240, 0]);
   "ROLL_State".M[77, 1] := #r;
   // PB16, STEP 5 network 16
   #r := ((((NOT "ROLL_IO".Input[12, 1]) AND ("ROLL_IO".Input[11, 1] OR "ROLL_IO".Input[11, 2] OR "ROLL_IO".Input[11, 3] OR "ROLL_IO".Input[11, 4] OR "ROLL_IO".Input[119, 6] OR "ROLL_IO".Input[119, 7] OR "ROLL_IO".Input[120, 0] OR "ROLL_IO".Input[120, 1])) OR (NOT "ROLL_IO".Input[12, 7])) AND ((NOT "ROLL_IO".Input[12, 7]) OR (NOT "ROLL_State".M[77, 1]) OR "ROLL_State".M[240, 0]) AND "ROLL_IO".Input[0, 1] AND "ROLL_IO".Input[11, 6] AND "ROLL_State".M[190, 6] AND "ROLL_State".M[23, 0]);
   "ROLL_State".M[77, 2] := #r;
   // PB16, STEP 5 network 17
   #r := (((NOT "ROLL_State".M[6, 0]) AND (NOT "ROLL_State".M[6, 2]) AND ("ROLL_IO".Input[11, 1] OR "ROLL_IO".Input[11, 2] OR "ROLL_IO".Input[11, 3] OR "ROLL_IO".Input[11, 4] OR "ROLL_IO".Input[119, 6] OR "ROLL_IO".Input[119, 7] OR "ROLL_IO".Input[120, 0])) OR "ROLL_IO".Input[11, 4]);
   "ROLL_State".M[76, 4] := #r;
   // PB16, STEP 5 network 18
   #r := ((NOT "ROLL_State".M[190, 5]) AND "ROLL_State".M[190, 6] AND "ROLL_State".M[23, 0] AND "ROLL_State".M[76, 4] AND "ROLL_State".M[77, 2]);
   "ROLL_State".M[76, 5] := #r;
   // PB16, STEP 5 network 19
   #r := ((((NOT "ROLL_State".M[190, 6]) AND "ROLL_State".M[190, 5] AND "ROLL_State".M[23, 0]) OR "ROLL_State".M[74, 0]) AND (("ROLL_IO".Input[124, 2] AND "ROLL_IO".Input[124, 5]) OR "ROLL_State".M[0, 4]) AND "ROLL_IO".Input[11, 0] AND "ROLL_State".M[63, 1]);
   "ROLL_State".M[76, 6] := #r;
   // PB16, STEP 5 network 20
   #r := (((((NOT "ROLL_IO".Input[12, 1]) OR (NOT "ROLL_IO".Input[12, 7])) AND "ROLL_State".M[76, 6]) OR "ROLL_State".M[76, 5]) AND "ROLL_IO".Input[0, 1] AND "ROLL_IO".Input[11, 6]);
   "ROLL_State".M[77, 0] := #r;
   // PB16, STEP 5 network 21
   #r := (((NOT "ROLL_IO".Input[11, 0]) AND (NOT "ROLL_IO".Input[12, 5]) AND "ROLL_State".M[190, 5]) OR ((NOT "ROLL_IO".Input[12, 1]) AND "ROLL_IO".Input[11, 0] AND "ROLL_State".M[190, 6]));
   "ROLL_State".M[240, 0] := #r;
   // PB16, STEP 5 network 22
   #r := ((NOT "ROLL_IO".Input[12, 1]) AND ("ROLL_IO".Input[11, 1] OR "ROLL_IO".Input[11, 2] OR "ROLL_IO".Input[11, 3] OR "ROLL_IO".Input[11, 4] OR "ROLL_IO".Input[119, 6] OR "ROLL_IO".Input[119, 7] OR "ROLL_IO".Input[120, 0]));
   "ROLL_State".M[240, 1] := #r;
   // PB16, STEP 5 network 23
   #r := ((NOT "ROLL_IO".Input[12, 1]) AND "ROLL_IO".Input[11, 0]);
   "ROLL_State".M[240, 2] := #r;
   // PB16, STEP 5 network 24
   #r := ((("ROLL_State".M[240, 1] OR "ROLL_State".M[240, 2]) AND "ROLL_State".M[77, 0]) OR ("ROLL_State".M[240, 0] AND "ROLL_State".M[76, 2]));
   "ROLL_State".M[76, 7] := #r;
   // PB16, STEP 5 network 25
   #r := ((NOT "ROLL_IO".Output[113, 3]) AND (NOT "ROLL_State".M[70, 2]) AND (NOT "ROLL_State".M[70, 3]) AND "ROLL_IO".Input[0, 1] AND "ROLL_IO".Input[11, 0] AND "ROLL_IO".Input[12, 1] AND "ROLL_IO".Input[12, 7] AND "ROLL_IO".Input[124, 5]);
   "ROLL_State".M[77, 3] := #r;
   // PB16, STEP 5 network 26
   #r := ((NOT "ROLL_State".M[77, 6]) AND (((NOT "ROLL_State".M[190, 6]) AND "ROLL_State".M[190, 5] AND "ROLL_State".M[22, 0]) OR "ROLL_State".M[74, 0]) AND "ROLL_IO".Output[113, 2] AND "ROLL_State".M[77, 3]);
   "ROLL_State".M[77, 4] := #r;
   // PB16, STEP 5 network 27
   #r := ((NOT "ROLL_State".M[190, 5]) AND (NOT "ROLL_State".M[77, 4]) AND "ROLL_State".M[190, 6] AND "ROLL_State".M[22, 0] AND "ROLL_State".M[77, 3]);
   "ROLL_State".M[77, 6] := #r;
   // PB16, STEP 5 network 28
   #r := ((NOT "ROLL_IO".Input[124, 5]) AND (NOT "ROLL_State".M[70, 3]) AND (((NOT "ROLL_IO".Input[124, 4]) AND "ROLL_State".M[20, 2] AND "ROLL_State".M[74, 0]) OR ((NOT "ROLL_State".M[190, 5]) AND "ROLL_IO".Input[0, 1] AND "ROLL_State".M[190, 6] AND "ROLL_State".M[22, 1])) AND "ROLL_IO".Input[124, 1]);
   "ROLL_State".M[77, 7] := #r;
   // PB16, STEP 5 network 29
   #r := ((NOT "ROLL_IO".Input[124, 4]) AND (NOT "ROLL_State".M[70, 3]) AND (((NOT "ROLL_State".M[15, 1]) AND "ROLL_State".M[20, 1] AND "ROLL_State".M[74, 0]) OR ((NOT "ROLL_State".M[190, 6]) AND "ROLL_IO".Input[0, 1] AND "ROLL_State".M[190, 5] AND "ROLL_State".M[22, 1])) AND "ROLL_IO".Input[124, 1]);
   "ROLL_State".M[78, 0] := #r;
   // PB16, STEP 5 network 30
   #r := ((("ROLL_State".M[22, 3] OR "ROLL_State".M[22, 4]) AND "ROLL_IO".Input[0, 1] AND "ROLL_State".M[190, 6]) OR ("ROLL_IO".Input[123, 5] AND "ROLL_State".M[74, 0]));
   IF #r THEN
       "ROLL_State".M[78, 4] := TRUE;
   END_IF;
   #r := (((NOT "ROLL_IO".Output[113, 3]) AND (NOT "ROLL_IO".Input[123, 4]) AND "ROLL_State".M[74, 0]) OR ((NOT "ROLL_IO".Output[113, 3]) AND "ROLL_IO".Input[0, 1] AND "ROLL_State".M[190, 5] AND "ROLL_State".M[22, 3]) OR (NOT "ROLL_IO".Input[0, 1]));
   IF #r THEN
       "ROLL_State".M[78, 4] := FALSE;
   END_IF;
   // PB16, STEP 5 network 31
   #r := ((NOT "ROLL_IO".Input[123, 5]) AND (NOT "ROLL_IO".Input[123, 6]) AND (NOT "ROLL_State".M[16, 0]) AND (NOT "ROLL_State".M[16, 4]) AND (NOT "ROLL_State".M[9, 1]) AND ((NOT "ROLL_IO".Input[123, 4]) OR "ROLL_State".M[190, 1]));
   "ROLL_State".M[78, 5] := #r;
   // PB16, STEP 5 network 32
   #r := (((NOT "ROLL_IO".Input[124, 2]) AND (NOT "ROLL_State".M[190, 5]) AND (NOT "ROLL_State".M[70, 3]) AND "ROLL_IO".Input[0, 1] AND "ROLL_IO".Input[124, 1] AND "ROLL_IO".Input[124, 4] AND "ROLL_State".M[190, 6] AND "ROLL_State".M[22, 4]) OR ("ROLL_State".M[70, 2] AND "ROLL_State".M[74, 0]));
   IF #r THEN
       "ROLL_State".M[78, 6] := TRUE;
   END_IF;
   #r := (((NOT "ROLL_State".M[70, 2]) AND ((NOT "ROLL_IO".Input[124, 1]) OR (NOT "ROLL_IO".Input[124, 4])) AND "ROLL_State".M[20, 2] AND "ROLL_State".M[74, 0]) OR ((NOT "ROLL_State".M[70, 2]) AND "ROLL_IO".Input[0, 1] AND "ROLL_State".M[190, 5] AND "ROLL_State".M[22, 4]) OR ((NOT "ROLL_State".M[70, 2]) AND "ROLL_State".M[20, 1] AND "ROLL_State".M[74, 0]) OR (NOT "ROLL_IO".Input[0, 1]) OR "ROLL_State".M[70, 0]);
   IF #r THEN
       "ROLL_State".M[78, 6] := FALSE;
   END_IF;
   // PB16, STEP 5 network 33
   #r := (((NOT "ROLL_State".M[70, 2]) AND (("ROLL_IO".Input[124, 5] AND "ROLL_State".M[20, 2]) OR "ROLL_State".M[20, 1]) AND "ROLL_State".M[74, 0]) OR ((NOT "ROLL_State".M[70, 2]) AND "ROLL_IO".Input[0, 1] AND "ROLL_State".M[190, 5] AND "ROLL_State".M[22, 4]));
   IF #r THEN
       "ROLL_State".M[78, 7] := TRUE;
   END_IF;
   #r := ((NOT "ROLL_IO".Input[0, 1]) OR "ROLL_State".M[70, 0] OR "ROLL_State".M[78, 6]);
   IF #r THEN
       "ROLL_State".M[78, 7] := FALSE;
   END_IF;
   // PB16, STEP 5 network 34
   RETURN;
END_FUNCTION

FUNCTION "ROLL_PB17" : Void   // FC25, SCL
{ S7_Optimized_Access := 'TRUE' }
VERSION : 0.1
// stored: AutoNumber true, IsIECCheckEnabled false, SetENOAutomatically false, UDAEnableTagReadback false
   VAR_TEMP
      r : Bool;
      a1 : Word;
      a2 : Word;
      activeDataBlock : Int;
      comparisonResults : Array[0..0] of Bool;
   END_VAR
BEGIN

